  movel([0.238520, -0.777638, -2.781210, -1.153541, 1.570796, 1.809316],accel_mss,speed_ms,0,blend_radius_m)
  movel([0.239014, -0.778562, -2.781058, -1.152769, 1.570796, 1.809811],accel_mss,speed_ms,0,blend_radius_m)
  movel([0.239003, -0.779791, -2.780855, -1.151743, 1.570796, 1.809799],accel_mss,speed_ms,0,blend_radius_m)
  movel([0.238262, -0.781308, -2.780604, -1.150477, 1.570796, 1.809059],accel_mss,speed_ms,0,blend_radius_m)
  movel([0.237067, -0.782563, -2.780395, -1.149431, 1.570796, 1.807864],accel_mss,speed_ms,0,blend_radius_m)
  movel([0.235771, -0.783294, -2.780273, -1.148822, 1.570796, 1.806567],accel_mss,speed_ms,0,blend_radius_m)
  movel([0.234495, -0.783612, -2.780219, -1.148557, 1.570796, 1.805291],accel_mss,speed_ms,0,blend_radius_m)
  movel([0.233364, -0.783640, -2.780215, -1.148534, 1.570796, 1.804160],accel_mss,speed_ms,0,blend_radius_m)
  movel([0.227228, -0.782889, -2.780340, -1.149160, 1.570796, 1.798025],accel_mss,speed_ms,0,blend_radius_m)
  movel([0.221349, -0.781729, -2.780534, -1.150126, 1.570796, 1.792145],accel_mss,speed_ms,0,blend_radius_m)
  movel([0.215730, -0.780164, -2.780794, -1.151432, 1.570796, 1.786526],accel_mss,speed_ms,0,blend_radius_m)
  movel([0.210389, -0.778185, -2.781120, -1.153084, 1.570796, 1.781185],accel_mss,speed_ms,0,blend_radius_m)
  movel([0.208538, -0.777277, -2.781269, -1.153843, 1.570796, 1.779334],accel_mss,speed_ms,0,blend_radius_m)
  movel([0.207075, -0.775893, -2.781496, -1.155000, 1.570796, 1.777871],accel_mss,speed_ms,0,blend_radius_m)
  movel([0.206532, -0.774726, -2.781686, -1.155977, 1.570796, 1.777328],accel_mss,speed_ms,0,blend_radius_m)
  movel([0.206197, -0.773361, -2.781908, -1.157121, 1.570796, 1.776993],accel_mss,speed_ms,0,blend_radius_m)
  movel([0.205895, -0.770284, -2.782404, -1.159701, 1.570796, 1.776692],accel_mss,speed_ms,0,blend_radius_m)
  movel([0.206072, -0.758256, -2.784298, -1.169835, 1.570796, 1.776868],accel_mss,speed_ms,0,blend_radius_m)
  movel([0.205767, -0.755116, -2.784781, -1.172493, 1.570796, 1.776563],accel_mss,speed_ms,0,blend_radius_m)
  movel([0.205061, -0.752630, -2.785159, -1.174600, 1.570796, 1.775857],accel_mss,speed_ms,0,blend_radius_m)
  movel([0.204513, -0.751748, -2.785293, -1.175348, 1.570796, 1.775309],accel_mss,speed_ms,0,blend_radius_m)
  movel([0.203813, -0.751162, -2.785382, -1.175845, 1.570796, 1.774609],accel_mss,speed_ms,0,blend_radius_m)
  movel([0.202946, -0.750924, -2.785418, -1.176048, 1.570796, 1.773742],accel_mss,speed_ms,0,blend_radius_m)
  movel([0.201896, -0.751069, -2.785396, -1.175924, 1.570796, 1.772693],accel_mss,speed_ms,0,blend_radius_m)
  movel([0.199844, -0.751927, -2.785266, -1.175196, 1.570796, 1.770640],accel_mss,speed_ms,0,blend_radius_m)
  movel([0.198900, -0.752216, -2.785222, -1.174950, 1.570796, 1.769696],accel_mss,speed_ms,0,blend_radius_m)
  movel([0.198186, -0.752114, -2.785238, -1.175037, 1.570796, 1.768982],accel_mss,speed_ms,0,blend_radius_m)
  movel([0.197823, -0.751113, -2.785389, -1.175887, 1.570796, 1.768619],accel_mss,speed_ms,0,blend_radius_m)
  movel([0.198037, -0.749591, -2.785618, -1.177180, 1.570796, 1.768834],accel_mss,speed_ms,0,blend_radius_m)
  movel([0.198952, -0.744572, -2.786366, -1.181452, 1.570796, 1.769748],accel_mss,speed_ms,0,blend_radius_m)
  movel([0.199542, -0.739772, -2.787069, -1.185548, 1.570796, 1.770338],accel_mss,speed_ms,0,blend_radius_m)
  movel([0.199909, -0.730710, -2.788367, -1.193312, 1.570796, 1.770705],accel_mss,speed_ms,0,blend_radius_m)
  movel([0.199495, -0.722125, -2.789560, -1.200704, 1.570796, 1.770291],accel_mss,speed_ms,0,blend_radius_m)
  movel([0.198653, -0.713738, -2.790692, -1.207959, 1.570796, 1.769449],accel_mss,speed_ms,0,blend_radius_m)
  speed_ms = 0.005
  movel([0.198653, -0.707172, -2.784094, -1.221123, 1.570796, 1.769449],accel_mss,speed_ms,0,blend_radius_m)
  speed_ms = 0.040
  movel([0.192703, -0.724050, -2.781792, -1.206547, 1.570796, 1.763499],accel_mss,speed_ms,0,blend_radius_m)
  speed_ms = 0.005
  movel([0.192703, -0.730831, -2.788350, -1.193208, 1.570796, 1.763499],accel_mss,speed_ms,0,blend_radius_m)
  speed_ms = 0.025
  movel([0.189482, -0.741949, -2.786751, -1.183689, 1.570796, 1.760279],accel_mss,speed_ms,0,blend_radius_m)
  movel([0.187584, -0.747603, -2.785916, -1.178870, 1.570796, 1.758381],accel_mss,speed_ms,0,blend_radius_m)
  movel([0.185510, -0.753297, -2.785058, -1.174034, 1.570796, 1.756306],accel_mss,speed_ms,0,blend_radius_m)
  movel([0.183050, -0.752490, -2.785181, -1.174719, 1.570796, 1.753846],accel_mss,speed_ms,0,blend_radius_m)
  movel([0.182585, -0.752423, -2.785191, -1.174775, 1.570796, 1.753381],accel_mss,speed_ms,0,blend_radius_m)
  movel([0.182001, -0.752685, -2.785151, -1.174553, 1.570796, 1.752798],accel_mss,speed_ms,0,blend_radius_m)
  movel([0.181431, -0.753357, -2.785049, -1.173983, 1.570796, 1.752227],accel_mss,speed_ms,0,blend_radius_m)
  movel([0.181021, -0.754135, -2.784931, -1.173324, 1.570796, 1.751817],accel_mss,speed_ms,0,blend_radius_m)
  movel([0.178486, -0.758934, -2.784193, -1.169262, 1.570796, 1.749283],accel_mss,speed_ms,0,blend_radius_m)
  movel([0.175445, -0.763691, -2.783451, -1.165247, 1.570796, 1.746242],accel_mss,speed_ms,0,blend_radius_m)
  movel([0.174614, -0.764748, -2.783285, -1.164356, 1.570796, 1.745410],accel_mss,speed_ms,0,blend_radius_m)
  movel([0.173739, -0.765391, -2.783183, -1.163814, 1.570796, 1.744535],accel_mss,speed_ms,0,blend_radius_m)
  movel([0.173247, -0.765240, -2.783207, -1.163942, 1.570796, 1.744044],accel_mss,speed_ms,0,blend_radius_m)
  movel([0.173079, -0.764663, -2.783298, -1.164428, 1.570796, 1.743875],accel_mss,speed_ms,0,blend_radius_m)
  movel([0.172930, -0.760434, -2.783961, -1.167994, 1.570796, 1.743726],accel_mss,speed_ms,0,blend_radius_m)
  movel([0.173553, -0.755646, -2.784700, -1.172043, 1.570796, 1.744349],accel_mss,speed_ms,0,blend_radius_m)
  speed_ms = 0.005
  movel([0.173553, -0.748568, -2.778205, -1.185616, 1.570796, 1.744349],accel_mss,speed_ms,0,blend_radius_m)
  speed_ms = 0.040
  movel([0.180746, -0.753780, -2.777404, -1.181204, 1.570796, 1.751543],accel_mss,speed_ms,0,blend_radius_m)
  speed_ms = 0.005
  movel([0.180746, -0.760919, -2.783885, -1.167585, 1.570796, 1.751543],accel_mss,speed_ms,0,blend_radius_m)
  speed_ms = 0.025
  movel([0.179875, -0.767925, -2.782781, -1.161683, 1.570796, 1.750672],accel_mss,speed_ms,0,blend_radius_m)
  movel([0.179084, -0.771629, -2.782188, -1.158572, 1.570796, 1.749880],accel_mss,speed_ms,0,blend_radius_m)
  movel([0.176839, -0.779327, -2.780932, -1.152130, 1.570796, 1.747635],accel_mss,speed_ms,0,blend_radius_m)
  movel([0.175396, -0.783288, -2.780274, -1.148827, 1.570796, 1.746192],accel_mss,speed_ms,0,blend_radius_m)
  movel([0.171908, -0.791341, -2.778911, -1.142138, 1.570796, 1.742704],accel_mss,speed_ms,0,blend_radius_m)
  movel([0.172377, -0.788931, -2.779322, -1.144136, 1.570796, 1.743174],accel_mss,speed_ms,0,blend_radius_m)
  movel([0.172203, -0.786949, -2.779658, -1.145782, 1.570796, 1.742999],accel_mss,speed_ms,0,blend_radius_m)
  movel([0.171413, -0.785526, -2.779898, -1.146964, 1.570796, 1.742209],accel_mss,speed_ms,0,blend_radius_m)
  movel([0.170034, -0.784796, -2.780021, -1.147572, 1.570796, 1.740831],accel_mss,speed_ms,0,blend_radius_m)
  speed_ms = 0.005
  movel([0.170034, -0.777395, -2.773605, -1.161389, 1.570796, 1.740831],accel_mss,speed_ms,0,blend_radius_m)
  speed_ms = 0.040
  movel([0.144449, -0.795994, -2.770410, -1.145985, 1.570796, 1.715246],accel_mss,speed_ms,0,blend_radius_m)
  speed_ms = 0.005
  movel([0.144449, -0.803590, -2.776772, -1.132027, 1.570796, 1.715246],accel_mss,speed_ms,0,blend_radius_m)
  speed_ms = 0.025
  movel([0.140306, -0.809331, -2.775742, -1.127316, 1.570796, 1.711102],accel_mss,speed_ms,0,blend_radius_m)
  movel([0.135816, -0.814795, -2.774745, -1.122849, 1.570796, 1.706612],accel_mss,speed_ms,0,blend_radius_m)
  movel([0.131062, -0.819901, -2.773799, -1.118689, 1.570796, 1.701858],accel_mss,speed_ms,0,blend_radius_m)
  movel([0.126121, -0.824563, -2.772923, -1.114904, 1.570796, 1.696917],accel_mss,speed_ms,0,blend_radius_m)
  movel([0.127219, -0.822105, -2.773386, -1.116898, 1.570796, 1.698016],accel_mss,speed_ms,0,blend_radius_m)
  movel([0.127994, -0.819853, -2.773808, -1.118728, 1.570796, 1.698790],accel_mss,speed_ms,0,blend_radius_m)
  movel([0.128392, -0.818004, -2.774152, -1.120233, 1.570796, 1.699188],accel_mss,speed_ms,0,blend_radius_m)
  movel([0.128362, -0.816754, -2.774384, -1.121251, 1.570796, 1.699159],accel_mss,speed_ms,0,blend_radius_m)
  movel([0.127847, -0.816316, -2.774465, -1.121608, 1.570796, 1.698643],accel_mss,speed_ms,0,blend_radius_m)
  movel([0.127395, -0.816460, -2.774438, -1.121491, 1.570796, 1.698191],accel_mss,speed_ms,0,blend_radius_m)
  movel([0.126795, -0.816881, -2.774360, -1.121147, 1.570796, 1.697592],accel_mss,speed_ms,0,blend_radius_m)
  movel([0.125163, -0.818650, -2.774032, -1.119707, 1.570796, 1.695960],accel_mss,speed_ms,0,blend_radius_m)
  movel([0.121164, -0.824312, -2.772970, -1.115107, 1.570796, 1.691961],accel_mss,speed_ms,0,blend_radius_m)
  movel([0.119283, -0.826786, -2.772500, -1.113103, 1.570796, 1.690079],accel_mss,speed_ms,0,blend_radius_m)
  movel([0.115192, -0.831505, -2.771595, -1.109289, 1.570796, 1.685989],accel_mss,speed_ms,0,blend_radius_m)
  movel([0.113032, -0.833691, -2.771171, -1.107526, 1.570796, 1.683829],accel_mss,speed_ms,0,blend_radius_m)
  movel([0.110826, -0.835714, -2.770777, -1.105898, 1.570796, 1.681622],accel_mss,speed_ms,0,blend_radius_m)
  movel([0.108596, -0.837553, -2.770416, -1.104420, 1.570796, 1.679392],accel_mss,speed_ms,0,blend_radius_m)
  movel([0.106371, -0.839163, -2.770099, -1.103127, 1.570796, 1.677167],accel_mss,speed_ms,0,blend_radius_m)
  movel([0.108926, -0.835167, -2.770884, -1.106338, 1.570796, 1.679722],accel_mss,speed_ms,0,blend_radius_m)
  movel([0.111408, -0.831132, -2.771667, -1.109590, 1.570796, 1.682204],accel_mss,speed_ms,0,blend_radius_m)
  movel([0.112472, -0.828577, -2.772158, -1.111654, 1.570796, 1.683268],accel_mss,speed_ms,0,blend_radius_m)
  movel([0.112976, -0.826234, -2.772605, -1.113550, 1.570796, 1.683773],accel_mss,speed_ms,0,blend_radius_m)
  movel([0.112833, -0.825536, -2.772738, -1.114115, 1.570796, 1.683630],accel_mss,speed_ms,0,blend_radius_m)
  movel([0.112322, -0.825368, -2.772770, -1.114251, 1.570796, 1.683118],accel_mss,speed_ms,0,blend_radius_m)
  movel([0.111378, -0.825886, -2.772672, -1.113832, 1.570796, 1.682174],accel_mss,speed_ms,0,blend_radius_m)
  movel([0.109924, -0.827249, -2.772412, -1.112728, 1.570796, 1.680720],accel_mss,speed_ms,0,blend_radius_m)
  movel([0.102400, -0.835431, -2.770832, -1.106126, 1.570796, 1.673197],accel_mss,speed_ms,0,blend_radius_m)
  movel([0.098589, -0.839089, -2.770114, -1.103186, 1.570796, 1.669385],accel_mss,speed_ms,0,blend_radius_m)
  movel([0.096654, -0.840643, -2.769806, -1.101939, 1.570796, 1.667451],accel_mss,speed_ms,0,blend_radius_m)
  movel([0.094689, -0.841956, -2.769545, -1.100887, 1.570796, 1.665485],accel_mss,speed_ms,0,blend_radius_m)
  speed_ms = 0.005
  movel([0.094689, -0.834001, -2.763299, -1.115089, 1.570796, 1.665485],accel_mss,speed_ms,0,blend_radius_m)
  speed_ms = 0.040
  movel([0.128026, -0.781141, -2.772976, -1.158272, 1.570796, 1.698822],accel_mss,speed_ms,0,blend_radius_m)
  speed_ms = 0.005
  movel([0.128026, -0.788583, -2.779381, -1.144425, 1.570796, 1.698822],accel_mss,speed_ms,0,blend_radius_m)
  speed_ms = 0.025
  movel([0.127894, -0.785887, -2.779837, -1.146664, 1.570796, 1.698691],accel_mss,speed_ms,0,blend_radius_m)
  movel([0.128371, -0.782803, -2.780355, -1.149231, 1.570796, 1.699168],accel_mss,speed_ms,0,blend_radius_m)
  movel([0.129395, -0.779405, -2.780919, -1.152065, 1.570796, 1.700191],accel_mss,speed_ms,0,blend_radius_m)
  movel([0.130900, -0.775786, -2.781513, -1.155090, 1.570796, 1.701697],accel_mss,speed_ms,0,blend_radius_m)
  movel([0.132838, -0.772016, -2.782125, -1.158247, 1.570796, 1.703635],accel_mss,speed_ms,0,blend_radius_m)
  movel([0.135137, -0.768197, -2.782738, -1.161454, 1.570796, 1.705933],accel_mss,speed_ms,0,blend_radius_m)
  movel([0.137743, -0.764400, -2.783340, -1.164649, 1.570796, 1.708540],accel_mss,speed_ms,0,blend_radius_m)
  movel([0.140583, -0.760728, -2.783915, -1.167746, 1.570796, 1.711379],accel_mss,speed_ms,0,blend_radius_m)
  movel([0.144308, -0.756402, -2.784584, -1.171403, 1.570796, 1.715105],accel_mss,speed_ms,0,blend_radius_m)
  movel([0.151976, -0.747852, -2.785879, -1.178659, 1.570796, 1.722772],accel_mss,speed_ms,0,blend_radius_m)
  movel([0.155648, -0.743371, -2.786543, -1.182475, 1.570796, 1.726445],accel_mss,speed_ms,0,blend_radius_m)
  movel([0.158985, -0.738544, -2.787247, -1.186598, 1.570796, 1.729782],accel_mss,speed_ms,0,blend_radius_m)
  movel([0.160417, -0.736070, -2.787604, -1.188715, 1.570796, 1.731214],accel_mss,speed_ms,0,blend_radius_m)
  movel([0.161621, -0.733642, -2.787951, -1.190796, 1.570796, 1.732417],accel_mss,speed_ms,0,blend_radius_m)
  movel([0.162542, -0.731323, -2.788280, -1.192786, 1.570796, 1.733339],accel_mss,speed_ms,0,blend_radius_m)
  movel([0.163134, -0.729175, -2.788583, -1.194631, 1.570796, 1.733930],accel_mss,speed_ms,0,blend_radius_m)
  movel([0.163330, -0.727280, -2.788848, -1.196261, 1.570796, 1.734126],accel_mss,speed_ms,0,blend_radius_m)
  movel([0.163076, -0.725704, -2.789067, -1.197618, 1.570796, 1.733872],accel_mss,speed_ms,0,blend_radius_m)
  speed_ms = 0.005
  movel([0.163076, -0.718987, -2.782497, -1.210906, 1.570796, 1.733872],accel_mss,speed_ms,0,blend_radius_m)
  speed_ms = 0.040
  movel([0.160050, -0.707154, -2.784096, -1.221139, 1.570796, 1.730846],accel_mss,speed_ms,0,blend_radius_m)
  speed_ms = 0.005
  movel([0.160050, -0.713719, -2.790695, -1.207975, 1.570796, 1.730846],accel_mss,speed_ms,0,blend_radius_m)
  speed_ms = 0.025
  movel([0.157424, -0.725682, -2.789070, -1.197637, 1.570796, 1.728221],accel_mss,speed_ms,0,blend_radius_m)
  movel([0.156311, -0.728566, -2.788668, -1.195155, 1.570796, 1.727108],accel_mss,speed_ms,0,blend_radius_m)
  movel([0.154500, -0.731547, -2.788249, -1.192593, 1.570796, 1.725296],accel_mss,speed_ms,0,blend_radius_m)
  movel([0.152223, -0.734414, -2.787841, -1.190134, 1.570796, 1.723019],accel_mss,speed_ms,0,blend_radius_m)
  movel([0.144460, -0.743032, -2.786593, -1.182764, 1.570796, 1.715257],accel_mss,speed_ms,0,blend_radius_m)
  movel([0.141887, -0.746260, -2.786116, -1.180013, 1.570796, 1.712683],accel_mss,speed_ms,0,blend_radius_m)
  movel([0.139486, -0.749568, -2.785622, -1.177199, 1.570796, 1.710282],accel_mss,speed_ms,0,blend_radius_m)
  movel([0.137275, -0.752916, -2.785116, -1.174357, 1.570796, 1.708071],accel_mss,speed_ms,0,blend_radius_m)
  movel([0.135464, -0.756183, -2.784617, -1.171588, 1.570796, 1.706261],accel_mss,speed_ms,0,blend_radius_m)
  movel([0.133979, -0.759398, -2.784121, -1.168869, 1.570796, 1.704776],accel_mss,speed_ms,0,blend_radius_m)
  movel([0.132528, -0.762585, -2.783625, -1.166179, 1.570796, 1.703325],accel_mss,speed_ms,0,blend_radius_m)
  movel([0.130825, -0.765773, -2.783123, -1.163493, 1.570796, 1.701621],accel_mss,speed_ms,0,blend_radius_m)
  movel([0.128528, -0.761127, -2.783853, -1.167409, 1.570796, 1.699324],accel_mss,speed_ms,0,blend_radius_m)
  movel([0.128585, -0.759365, -2.784127, -1.168898, 1.570796, 1.699381],accel_mss,speed_ms,0,blend_radius_m)
  movel([0.128955, -0.757448, -2.784423, -1.170518, 1.570796, 1.699752],accel_mss,speed_ms,0,blend_radius_m)
  movel([0.129638, -0.755372, -2.784742, -1.172275, 1.570796, 1.700435],accel_mss,speed_ms,0,blend_radius_m)
  movel([0.130651, -0.753118, -2.785085, -1.174186, 1.570796, 1.701447],accel_mss,speed_ms,0,blend_radius_m)
  movel([0.132666, -0.749871, -2.785576, -1.176942, 1.570796, 1.703462],accel_mss,speed_ms,0,blend_radius_m)
  movel([0.135700, -0.745820, -2.786181, -1.180388, 1.570796, 1.706497],accel_mss,speed_ms,0,blend_radius_m)
  movel([0.143277, -0.736531, -2.787538, -1.188320, 1.570796, 1.714073],accel_mss,speed_ms,0,blend_radius_m)
  movel([0.147031, -0.731929, -2.788195, -1.192265, 1.570796, 1.717828],accel_mss,speed_ms,0,blend_radius_m)
  movel([0.150221, -0.727782, -2.788778, -1.195829, 1.570796, 1.721017],accel_mss,speed_ms,0,blend_radius_m)
  movel([0.152429, -0.724431, -2.789243, -1.198715, 1.570796, 1.723225],accel_mss,speed_ms,0,blend_radius_m)
  movel([0.153036, -0.723152, -2.789419, -1.199818, 1.570796, 1.723833],accel_mss,speed_ms,0,blend_radius_m)
  movel([0.153239, -0.722197, -2.789550, -1.200642, 1.570796, 1.724035],accel_mss,speed_ms,0,blend_radius_m)
  speed_ms = 0.005
  movel([0.153239, -0.715524, -2.782972, -1.213894, 1.570796, 1.724035],accel_mss,speed_ms,0,blend_radius_m)
  speed_ms = 0.040
  movel([0.137879, -0.720219, -2.782326, -1.209843, 1.570796, 1.708675],accel_mss,speed_ms,0,blend_radius_m)
  speed_ms = 0.005
  movel([0.137879, -0.726952, -2.788893, -1.196543, 1.570796, 1.708675],accel_mss,speed_ms,0,blend_radius_m)
  speed_ms = 0.025
  movel([0.136395, -0.727386, -2.788833, -1.196170, 1.570796, 1.707191],accel_mss,speed_ms,0,blend_radius_m)
  movel([0.135134, -0.727419, -2.788828, -1.196142, 1.570796, 1.705931],accel_mss,speed_ms,0,blend_radius_m)
  movel([0.133190, -0.726532, -2.788952, -1.196905, 1.570796, 1.703986],accel_mss,speed_ms,0,blend_radius_m)
  movel([0.131847, -0.724748, -2.789199, -1.198441, 1.570796, 1.702644],accel_mss,speed_ms,0,blend_radius_m)
  movel([0.130926, -0.722510, -2.789507, -1.200371, 1.570796, 1.701722],accel_mss,speed_ms,0,blend_radius_m)
  movel([0.130785, -0.721530, -2.789642, -1.201218, 1.570796, 1.701582],accel_mss,speed_ms,0,blend_radius_m)
  movel([0.131601, -0.719398, -2.789932, -1.203059, 1.570796, 1.702397],accel_mss,speed_ms,0,blend_radius_m)
  movel([0.134610, -0.713129, -2.790773, -1.208487, 1.570796, 1.705407],accel_mss,speed_ms,0,blend_radius_m)
  movel([0.140137, -0.700606, -2.792400, -1.219383, 1.570796, 1.710933],accel_mss,speed_ms,0,blend_radius_m)
  movel([0.142639, -0.694384, -2.793181, -1.224825, 1.570796, 1.713435],accel_mss,speed_ms,0,blend_radius_m)
  speed_ms = 0.005
  movel([0.142639, -0.688072, -2.786538, -1.237779, 1.570796, 1.713435],accel_mss,speed_ms,0,blend_radius_m)
  speed_ms = 0.040
  movel([0.132933, -0.695886, -2.785558, -1.230945, 1.570796, 1.703729],accel_mss,speed_ms,0,blend_radius_m)
  speed_ms = 0.005
  movel([0.132933, -0.702302, -2.792184, -1.217903, 1.570796, 1.703729],accel_mss,speed_ms,0,blend_radius_m)
  speed_ms = 0.025
  movel([0.131774, -0.705905, -2.791720, -1.214763, 1.570796, 1.702571],accel_mss,speed_ms,0,blend_radius_m)
  movel([0.130233, -0.709651, -2.791232, -1.211506, 1.570796, 1.701029],accel_mss,speed_ms,0,blend_radius_m)
  movel([0.128199, -0.713401, -2.790737, -1.208251, 1.570796, 1.698995],accel_mss,speed_ms,0,blend_radius_m)
  movel([0.126962, -0.715242, -2.790492, -1.206655, 1.570796, 1.697758],accel_mss,speed_ms,0,blend_radius_m)
  movel([0.124214, -0.718795, -2.790014, -1.203580, 1.570796, 1.695010],accel_mss,speed_ms,0,blend_radius_m)
  movel([0.123618, -0.720283, -2.789812, -1.202294, 1.570796, 1.694414],accel_mss,speed_ms,0,blend_radius_m)
  movel([0.120317, -0.731224, -2.788294, -1.192871, 1.570796, 1.691113],accel_mss,speed_ms,0,blend_radius_m)
  movel([0.120030, -0.732265, -2.788147, -1.191977, 1.570796, 1.690826],accel_mss,speed_ms,0,blend_radius_m)
  movel([0.120015, -0.733114, -2.788027, -1.191249, 1.570796, 1.690811],accel_mss,speed_ms,0,blend_radius_m)
  movel([0.120743, -0.733613, -2.787955, -1.190820, 1.570796, 1.691539],accel_mss,speed_ms,0,blend_radius_m)
  movel([0.121930, -0.733493, -2.787972, -1.190923, 1.570796, 1.692726],accel_mss,speed_ms,0,blend_radius_m)
  movel([0.125409, -0.732988, -2.788044, -1.191356, 1.570796, 1.696206],accel_mss,speed_ms,0,blend_radius_m)
  movel([0.128620, -0.732965, -2.788048, -1.191376, 1.570796, 1.699416],accel_mss,speed_ms,0,blend_radius_m)
  movel([0.131341, -0.733654, -2.787950, -1.190785, 1.570796, 1.702138],accel_mss,speed_ms,0,blend_radius_m)
  movel([0.133335, -0.735302, -2.787714, -1.189373, 1.570796, 1.704131],accel_mss,speed_ms,0,blend_radius_m)
  speed_ms = 0.005
  movel([0.133335, -0.728466, -2.781168, -1.202756, 1.570796, 1.704131],accel_mss,speed_ms,0,blend_radius_m)
  speed_ms = 0.040
  movel([0.124946, -0.756050, -2.777052, -1.179288, 1.570796, 1.695742],accel_mss,speed_ms,0,blend_radius_m)
  speed_ms = 0.005
  movel([0.124946, -0.763214, -2.783526, -1.165648, 1.570796, 1.695742],accel_mss,speed_ms,0,blend_radius_m)
  speed_ms = 0.025
  movel([0.124279, -0.763945, -2.783411, -1.165033, 1.570796, 1.695076],accel_mss,speed_ms,0,blend_radius_m)
  movel([0.123694, -0.764818, -2.783274, -1.164297, 1.570796, 1.694491],accel_mss,speed_ms,0,blend_radius_m)
  movel([0.121456, -0.769175, -2.782582, -1.160632, 1.570796, 1.692253],accel_mss,speed_ms,0,blend_radius_m)
  movel([0.121055, -0.769619, -2.782511, -1.160259, 1.570796, 1.691851],accel_mss,speed_ms,0,blend_radius_m)
  movel([0.120432, -0.769904, -2.782465, -1.160020, 1.570796, 1.691229],accel_mss,speed_ms,0,blend_radius_m)
  movel([0.119925, -0.769768, -2.782487, -1.160134, 1.570796, 1.690722],accel_mss,speed_ms,0,blend_radius_m)
  movel([0.119237, -0.768645, -2.782667, -1.161078, 1.570796, 1.690033],accel_mss,speed_ms,0,blend_radius_m)
  movel([0.118835, -0.765855, -2.783110, -1.163424, 1.570796, 1.689631],accel_mss,speed_ms,0,blend_radius_m)
  movel([0.119383, -0.762634, -2.783617, -1.166137, 1.570796, 1.690179],accel_mss,speed_ms,0,blend_radius_m)
  movel([0.120418, -0.759122, -2.784164, -1.169102, 1.570796, 1.691215],accel_mss,speed_ms,0,blend_radius_m)
  movel([0.121709, -0.755540, -2.784716, -1.172133, 1.570796, 1.692506],accel_mss,speed_ms,0,blend_radius_m)
  movel([0.123298, -0.751966, -2.785260, -1.175163, 1.570796, 1.694094],accel_mss,speed_ms,0,blend_radius_m)
  movel([0.125173, -0.748402, -2.785796, -1.178190, 1.570796, 1.695969],accel_mss,speed_ms,0,blend_radius_m)
  movel([0.127322, -0.744851, -2.786324, -1.181213, 1.570796, 1.698119],accel_mss,speed_ms,0,blend_radius_m)
  movel([0.129739, -0.741309, -2.786845, -1.184235, 1.570796, 1.700535],accel_mss,speed_ms,0,blend_radius_m)
  movel([0.132404, -0.737785, -2.787357, -1.187247, 1.570796, 1.703200],accel_mss,speed_ms,0,blend_radius_m)
  movel([0.135317, -0.734268, -2.787862, -1.190259, 1.570796, 1.706113],accel_mss,speed_ms,0,blend_radius_m)
  movel([0.138458, -0.730769, -2.788359, -1.193261, 1.570796, 1.709254],accel_mss,speed_ms,0,blend_radius_m)
  movel([0.142773, -0.725595, -2.789082, -1.197712, 1.570796, 1.713570],accel_mss,speed_ms,0,blend_radius_m)
  movel([0.147235, -0.719614, -2.789903, -1.202872, 1.570796, 1.718031],accel_mss,speed_ms,0,blend_radius_m)
  movel([0.152015, -0.712739, -2.790825, -1.208825, 1.570796, 1.722812],accel_mss,speed_ms,0,blend_radius_m)
  speed_ms = 0.005
  movel([0.152015, -0.706186, -2.784224, -1.221979, 1.570796, 1.722812],accel_mss,speed_ms,0,blend_radius_m)
  speed_ms = 0.040
  movel([0.147515, -0.708228, -2.783953, -1.220207, 1.570796, 1.718311],accel_mss,speed_ms,0,blend_radius_m)
  speed_ms = 0.005
  movel([0.147515, -0.714808, -2.790550, -1.207031, 1.570796, 1.718311],accel_mss,speed_ms,0,blend_radius_m)
  speed_ms = 0.025
  movel([0.150955, -0.705951, -2.791714, -1.214723, 1.570796, 1.721751],accel_mss,speed_ms,0,blend_radius_m)
  movel([0.154901, -0.696855, -2.792873, -1.222662, 1.570796, 1.725698],accel_mss,speed_ms,0,blend_radius_m)
  movel([0.157180, -0.692234, -2.793447, -1.226708, 1.570796, 1.727976],accel_mss,speed_ms,0,blend_radius_m)
  movel([0.159708, -0.687580, -2.794015, -1.230794, 1.570796, 1.730504],accel_mss,speed_ms,0,blend_radius_m)
  movel([0.162546, -0.682891, -2.794578, -1.234920, 1.570796, 1.733342],accel_mss,speed_ms,0,blend_radius_m)
  movel([0.165720, -0.678193, -2.795132, -1.239064, 1.570796, 1.736517],accel_mss,speed_ms,0,blend_radius_m)
  movel([0.174701, -0.666260, -2.796496, -1.249633, 1.570796, 1.745498],accel_mss,speed_ms,0,blend_radius_m)
  movel([0.178567, -0.660821, -2.797097, -1.254472, 1.570796, 1.749363],accel_mss,speed_ms,0,blend_radius_m)
  movel([0.180369, -0.658058, -2.797397, -1.256934, 1.570796, 1.751165],accel_mss,speed_ms,0,blend_radius_m)
  movel([0.181974, -0.655275, -2.797696, -1.259418, 1.570796, 1.752770],accel_mss,speed_ms,0,blend_radius_m)
  movel([0.185372, -0.647161, -2.798550, -1.266679, 1.570796, 1.756168],accel_mss,speed_ms,0,blend_radius_m)
  speed_ms = 0.005
  movel([0.185372, -0.641516, -2.791809, -1.279065, 1.570796, 1.756168],accel_mss,speed_ms,0,blend_radius_m)
  speed_ms = 0.040
  movel([0.193729, -0.622779, -2.793665, -1.295945, 1.570796, 1.764526],accel_mss,speed_ms,0,blend_radius_m)
  speed_ms = 0.005
  movel([0.193729, -0.628139, -2.800441, -1.283810, 1.570796, 1.764526],accel_mss,speed_ms,0,blend_radius_m)
  speed_ms = 0.025
  movel([0.196333, -0.621490, -2.801066, -1.289833, 1.570796, 1.767130],accel_mss,speed_ms,0,blend_radius_m)
  movel([0.198154, -0.618053, -2.801382, -1.292954, 1.570796, 1.768950],accel_mss,speed_ms,0,blend_radius_m)
  movel([0.200526, -0.614603, -2.801695, -1.296091, 1.570796, 1.771322],accel_mss,speed_ms,0,blend_radius_m)
  movel([0.202505, -0.612299, -2.801901, -1.298189, 1.570796, 1.773301],accel_mss,speed_ms,0,blend_radius_m)
  movel([0.204614, -0.610164, -2.802090, -1.300135, 1.570796, 1.775410],accel_mss,speed_ms,0,blend_radius_m)
  movel([0.209001, -0.606162, -2.802439, -1.303789, 1.570796, 1.779798],accel_mss,speed_ms,0,blend_radius_m)
  movel([0.212909, -0.602297, -2.802770, -1.307322, 1.570796, 1.783705],accel_mss,speed_ms,0,blend_radius_m)
  movel([0.215989, -0.598561, -2.803084, -1.310744, 1.570796, 1.786785],accel_mss,speed_ms,0,blend_radius_m)
  movel([0.221767, -0.590075, -2.803777, -1.318537, 1.570796, 1.792563],accel_mss,speed_ms,0,blend_radius_m)
  movel([0.223037, -0.588369, -2.803913, -1.320107, 1.570796, 1.793834],accel_mss,speed_ms,0,blend_radius_m)
  movel([0.224449, -0.586785, -2.804038, -1.321566, 1.570796, 1.795245],accel_mss,speed_ms,0,blend_radius_m)
  movel([0.227568, -0.583894, -2.804264, -1.324231, 1.570796, 1.798364],accel_mss,speed_ms,0,blend_radius_m)
  movel([0.233995, -0.578551, -2.804672, -1.329165, 1.570796, 1.804791],accel_mss,speed_ms,0,blend_radius_m)
  movel([0.240772, -0.572320, -2.805135, -1.334934, 1.570796, 1.811568],accel_mss,speed_ms,0,blend_radius_m)
  movel([0.244115, -0.568952, -2.805378, -1.338059, 1.570796, 1.814911],accel_mss,speed_ms,0,blend_radius_m)
  movel([0.247325, -0.565306, -2.805637, -1.341446, 1.570796, 1.818121],accel_mss,speed_ms,0,blend_radius_m)
  movel([0.249641, -0.562122, -2.805859, -1.344408, 1.570796, 1.820438],accel_mss,speed_ms,0,blend_radius_m)
  movel([0.251409, -0.558950, -2.806075, -1.347363, 1.570796, 1.822205],accel_mss,speed_ms,0,blend_radius_m)
  movel([0.252187, -0.556399, -2.806247, -1.349743, 1.570796, 1.822983],accel_mss,speed_ms,0,blend_radius_m)
  movel([0.252068, -0.555552, -2.806304, -1.350534, 1.570796, 1.822864],accel_mss,speed_ms,0,blend_radius_m)
  movel([0.251533, -0.555093, -2.806334, -1.350962, 1.570796, 1.822330],accel_mss,speed_ms,0,blend_radius_m)
  movel([0.249691, -0.555064, -2.806336, -1.350989, 1.570796, 1.820487],accel_mss,speed_ms,0,blend_radius_m)
  movel([0.247199, -0.555806, -2.806287, -1.350296, 1.570796, 1.817995],accel_mss,speed_ms,0,blend_radius_m)
  movel([0.244223, -0.557208, -2.806193, -1.348988, 1.570796, 1.815020],accel_mss,speed_ms,0,blend_radius_m)
  movel([0.240967, -0.559117, -2.806064, -1.347208, 1.570796, 1.811764],accel_mss,speed_ms,0,blend_radius_m)
  movel([0.237607, -0.561424, -2.805907, -1.345059, 1.570796, 1.808403],accel_mss,speed_ms,0,blend_radius_m)
  movel([0.234331, -0.563983, -2.805729, -1.342677, 1.570796, 1.805127],accel_mss,speed_ms,0,blend_radius_m)
  movel([0.231319, -0.566673, -2.805541, -1.340176, 1.570796, 1.802115],accel_mss,speed_ms,0,blend_radius_m)
  movel([0.228747, -0.569367, -2.805348, -1.337674, 1.570796, 1.799543],accel_mss,speed_ms,0,blend_radius_m)
  movel([0.225354, -0.573742, -2.805031, -1.333617, 1.570796, 1.796150],accel_mss,speed_ms,0,blend_radius_m)
  movel([0.216091, -0.586999, -2.804021, -1.321368, 1.570796, 1.786887],accel_mss,speed_ms,0,blend_radius_m)
  movel([0.209605, -0.595587, -2.803330, -1.313472, 1.570796, 1.780401],accel_mss,speed_ms,0,blend_radius_m)
  movel([0.203573, -0.602636, -2.802741, -1.307012, 1.570796, 1.774369],accel_mss,speed_ms,0,blend_radius_m)
  movel([0.200581, -0.606065, -2.802447, -1.303877, 1.570796, 1.771378],accel_mss,speed_ms,0,blend_radius_m)
  movel([0.197793, -0.609574, -2.802142, -1.300674, 1.570796, 1.768589],accel_mss,speed_ms,0,blend_radius_m)
  movel([0.195217, -0.613309, -2.801811, -1.297269, 1.570796, 1.766013],accel_mss,speed_ms,0,blend_radius_m)
  movel([0.192956, -0.617013, -2.801477, -1.293898, 1.570796, 1.763753],accel_mss,speed_ms,0,blend_radius_m)
  movel([0.190975, -0.620680, -2.801141, -1.290568, 1.570796, 1.761772],accel_mss,speed_ms,0,blend_radius_m)
  movel([0.189235, -0.624290, -2.800805, -1.287294, 1.570796, 1.760032],accel_mss,speed_ms,0,blend_radius_m)
  movel([0.186322, -0.631317, -2.800135, -1.280937, 1.570796, 1.757118],accel_mss,speed_ms,0,blend_radius_m)
  movel([0.183895, -0.638024, -2.799477, -1.274888, 1.570796, 1.754691],accel_mss,speed_ms,0,blend_radius_m)
  speed_ms = 0.005
  movel([0.183895, -0.632515, -2.792719, -1.287155, 1.570796, 1.754691],accel_mss,speed_ms,0,blend_radius_m)
  speed_ms = 0.040
  movel([0.176152, -0.639775, -2.791987, -1.280627, 1.570796, 1.746948],accel_mss,speed_ms,0,blend_radius_m)
  speed_ms = 0.005
  movel([0.176152, -0.645394, -2.798732, -1.268264, 1.570796, 1.746948],accel_mss,speed_ms,0,blend_radius_m)
  speed_ms = 0.025
  movel([0.180224, -0.634747, -2.799801, -1.277841, 1.570796, 1.751020],accel_mss,speed_ms,0,blend_radius_m)
  movel([0.182120, -0.630206, -2.800243, -1.281940, 1.570796, 1.752916],accel_mss,speed_ms,0,blend_radius_m)
  movel([0.183798, -0.625753, -2.800667, -1.285969, 1.570796, 1.754594],accel_mss,speed_ms,0,blend_radius_m)
  movel([0.184805, -0.622128, -2.801007, -1.289254, 1.570796, 1.755601],accel_mss,speed_ms,0,blend_radius_m)
  movel([0.185326, -0.618806, -2.801313, -1.292269, 1.570796, 1.756122],accel_mss,speed_ms,0,blend_radius_m)
  movel([0.185349, -0.615856, -2.801582, -1.294951, 1.570796, 1.756145],accel_mss,speed_ms,0,blend_radius_m)
  movel([0.184865, -0.613347, -2.801807, -1.297234, 1.570796, 1.755661],accel_mss,speed_ms,0,blend_radius_m)
  movel([0.186494, -0.611974, -2.801930, -1.298485, 1.570796, 1.757290],accel_mss,speed_ms,0,blend_radius_m)
  movel([0.188104, -0.610937, -2.802022, -1.299431, 1.570796, 1.758900],accel_mss,speed_ms,0,blend_radius_m)
  movel([0.191272, -0.609291, -2.802166, -1.300932, 1.570796, 1.762069],accel_mss,speed_ms,0,blend_radius_m)
  movel([0.194593, -0.607312, -2.802339, -1.302738, 1.570796, 1.765389],accel_mss,speed_ms,0,blend_radius_m)
  movel([0.196244, -0.605965, -2.802456, -1.303968, 1.570796, 1.767041],accel_mss,speed_ms,0,blend_radius_m)
  movel([0.197767, -0.604278, -2.802601, -1.305510, 1.570796, 1.768564],accel_mss,speed_ms,0,blend_radius_m)
  movel([0.214731, -0.582487, -2.804372, -1.325529, 1.570796, 1.785527],accel_mss,speed_ms,0,blend_radius_m)
  movel([0.214676, -0.580480, -2.804526, -1.327383, 1.570796, 1.785472],accel_mss,speed_ms,0,blend_radius_m)
  movel([0.213877, -0.579104, -2.804631, -1.328655, 1.570796, 1.784674],accel_mss,speed_ms,0,blend_radius_m)
  movel([0.212377, -0.578432, -2.804681, -1.329276, 1.570796, 1.783174],accel_mss,speed_ms,0,blend_radius_m)
  movel([0.210246, -0.578518, -2.804675, -1.329196, 1.570796, 1.781042],accel_mss,speed_ms,0,blend_radius_m)
  movel([0.214128, -0.575879, -2.804873, -1.331638, 1.570796, 1.784924],accel_mss,speed_ms,0,blend_radius_m)
  movel([0.217788, -0.573955, -2.805015, -1.333419, 1.570796, 1.788584],accel_mss,speed_ms,0,blend_radius_m)
  movel([0.221033, -0.572837, -2.805097, -1.334456, 1.570796, 1.791829],accel_mss,speed_ms,0,blend_radius_m)
  movel([0.223683, -0.572603, -2.805114, -1.334672, 1.570796, 1.794480],accel_mss,speed_ms,0,blend_radius_m)
  speed_ms = 0.005
  movel([0.223683, -0.568129, -2.798249, -1.346011, 1.570796, 1.794480],accel_mss,speed_ms,0,blend_radius_m)
  speed_ms = 0.040
  movel([0.226080, -0.558963, -2.798901, -1.354525, 1.570796, 1.796876],accel_mss,speed_ms,0,blend_radius_m)
  speed_ms = 0.005
  movel([0.226080, -0.563281, -2.805778, -1.343330, 1.570796, 1.796876],accel_mss,speed_ms,0,blend_radius_m)
  speed_ms = 0.025
  movel([0.228138, -0.557951, -2.806143, -1.348295, 1.570796, 1.798934],accel_mss,speed_ms,0,blend_radius_m)
  movel([0.229724, -0.553041, -2.806469, -1.352878, 1.570796, 1.800520],accel_mss,speed_ms,0,blend_radius_m)
  movel([0.230868, -0.548512, -2.806762, -1.357115, 1.570796, 1.801665],accel_mss,speed_ms,0,blend_radius_m)
  movel([0.231595, -0.544322, -2.807026, -1.361041, 1.570796, 1.802391],accel_mss,speed_ms,0,blend_radius_m)
  movel([0.231931, -0.540427, -2.807265, -1.364697, 1.570796, 1.802727],accel_mss,speed_ms,0,blend_radius_m)
  movel([0.231904, -0.536780, -2.807484, -1.368125, 1.570796, 1.802701],accel_mss,speed_ms,0,blend_radius_m)
  movel([0.230885, -0.530050, -2.807875, -1.374465, 1.570796, 1.801682],accel_mss,speed_ms,0,blend_radius_m)
  movel([0.224092, -0.548238, -2.806779, -1.357371, 1.570796, 1.794888],accel_mss,speed_ms,0,blend_radius_m)
  movel([0.224651, -0.546332, -2.806900, -1.359157, 1.570796, 1.795447],accel_mss,speed_ms,0,blend_radius_m)
  movel([0.224852, -0.544671, -2.807004, -1.360714, 1.570796, 1.795649],accel_mss,speed_ms,0,blend_radius_m)
  movel([0.224312, -0.542032, -2.807167, -1.363190, 1.570796, 1.795109],accel_mss,speed_ms,0,blend_radius_m)
  movel([0.222714, -0.540224, -2.807278, -1.364887, 1.570796, 1.793510],accel_mss,speed_ms,0,blend_radius_m)
  movel([0.220333, -0.539136, -2.807343, -1.365909, 1.570796, 1.791129],accel_mss,speed_ms,0,blend_radius_m)
  movel([0.217432, -0.538649, -2.807373, -1.366367, 1.570796, 1.788229],accel_mss,speed_ms,0,blend_radius_m)
  movel([0.214292, -0.538644, -2.807373, -1.366372, 1.570796, 1.785088],accel_mss,speed_ms,0,blend_radius_m)
  movel([0.208391, -0.539580, -2.807317, -1.365493, 1.570796, 1.779188],accel_mss,speed_ms,0,blend_radius_m)
  movel([0.211122, -0.543986, -2.807047, -1.361356, 1.570796, 1.781918],accel_mss,speed_ms,0,blend_radius_m)
  movel([0.211813, -0.546927, -2.806863, -1.358599, 1.570796, 1.782610],accel_mss,speed_ms,0,blend_radius_m)
  movel([0.211526, -0.550446, -2.806638, -1.355305, 1.570796, 1.782322],accel_mss,speed_ms,0,blend_radius_m)
  movel([0.209060, -0.551580, -2.806565, -1.354245, 1.570796, 1.779856],accel_mss,speed_ms,0,blend_radius_m)
  movel([0.206761, -0.552256, -2.806521, -1.353612, 1.570796, 1.777558],accel_mss,speed_ms,0,blend_radius_m)
  movel([0.202396, -0.552864, -2.806481, -1.353044, 1.570796, 1.773192],accel_mss,speed_ms,0,blend_radius_m)
  movel([0.197929, -0.553484, -2.806440, -1.352464, 1.570796, 1.768725],accel_mss,speed_ms,0,blend_radius_m)
  movel([0.195504, -0.554176, -2.806395, -1.351818, 1.570796, 1.766300],accel_mss,speed_ms,0,blend_radius_m)
  movel([0.192883, -0.555309, -2.806320, -1.350760, 1.570796, 1.763679],accel_mss,speed_ms,0,blend_radius_m)
  movel([0.190652, -0.560199, -2.805991, -1.346199, 1.570796, 1.761448],accel_mss,speed_ms,0,blend_radius_m)
  movel([0.189350, -0.564603, -2.805686, -1.342100, 1.570796, 1.760146],accel_mss,speed_ms,0,blend_radius_m)
  movel([0.185745, -0.566570, -2.805548, -1.340271, 1.570796, 1.756542],accel_mss,speed_ms,0,blend_radius_m)
  movel([0.182404, -0.567911, -2.805453, -1.339025, 1.570796, 1.753200],accel_mss,speed_ms,0,blend_radius_m)
  movel([0.179388, -0.568602, -2.805403, -1.338384, 1.570796, 1.750184],accel_mss,speed_ms,0,blend_radius_m)
  movel([0.176782, -0.568621, -2.805402, -1.338366, 1.570796, 1.747579],accel_mss,speed_ms,0,blend_radius_m)
  movel([0.176392, -0.569179, -2.805362, -1.337848, 1.570796, 1.747188],accel_mss,speed_ms,0,blend_radius_m)
  movel([0.173374, -0.575341, -2.804912, -1.332135, 1.570796, 1.744170],accel_mss,speed_ms,0,blend_radius_m)
  movel([0.169984, -0.582867, -2.804343, -1.325179, 1.570796, 1.740781],accel_mss,speed_ms,0,blend_radius_m)
  movel([0.168807, -0.586291, -2.804077, -1.322021, 1.570796, 1.739603],accel_mss,speed_ms,0,blend_radius_m)
  movel([0.168021, -0.589300, -2.803839, -1.319250, 1.570796, 1.738817],accel_mss,speed_ms,0,blend_radius_m)
  movel([0.167144, -0.595092, -2.803371, -1.313927, 1.570796, 1.737940],accel_mss,speed_ms,0,blend_radius_m)
  movel([0.158403, -0.593767, -2.803479, -1.315143, 1.570796, 1.729200],accel_mss,speed_ms,0,blend_radius_m)
  movel([0.157042, -0.597412, -2.803180, -1.311797, 1.570796, 1.727839],accel_mss,speed_ms,0,blend_radius_m)
  movel([0.155985, -0.600919, -2.802886, -1.308583, 1.570796, 1.726781],accel_mss,speed_ms,0,blend_radius_m)
  movel([0.154661, -0.607511, -2.802322, -1.302556, 1.570796, 1.725457],accel_mss,speed_ms,0,blend_radius_m)
  movel([0.154262, -0.613434, -2.801800, -1.297156, 1.570796, 1.725059],accel_mss,speed_ms,0,blend_radius_m)
  movel([0.154695, -0.620188, -2.801187, -1.291014, 1.570796, 1.725492],accel_mss,speed_ms,0,blend_radius_m)
  movel([0.154495, -0.621135, -2.801099, -1.290155, 1.570796, 1.725292],accel_mss,speed_ms,0,blend_radius_m)
  movel([0.154014, -0.622210, -2.800999, -1.289180, 1.570796, 1.724810],accel_mss,speed_ms,0,blend_radius_m)
  movel([0.152932, -0.623706, -2.800860, -1.287824, 1.570796, 1.723728],accel_mss,speed_ms,0,blend_radius_m)
  movel([0.144473, -0.632526, -2.800018, -1.279845, 1.570796, 1.715269],accel_mss,speed_ms,0,blend_radius_m)
  movel([0.140094, -0.636517, -2.799627, -1.276246, 1.570796, 1.710890],accel_mss,speed_ms,0,blend_radius_m)
  movel([0.138438, -0.637671, -2.799512, -1.275206, 1.570796, 1.709235],accel_mss,speed_ms,0,blend_radius_m)
  movel([0.137413, -0.637922, -2.799487, -1.274980, 1.570796, 1.708210],accel_mss,speed_ms,0,blend_radius_m)
  movel([0.141719, -0.639134, -2.799366, -1.273889, 1.570796, 1.712515],accel_mss,speed_ms,0,blend_radius_m)
  movel([0.144168, -0.639301, -2.799349, -1.273738, 1.570796, 1.714964],accel_mss,speed_ms,0,blend_radius_m)
  movel([0.146793, -0.639184, -2.799361, -1.273844, 1.570796, 1.717590],accel_mss,speed_ms,0,blend_radius_m)
  movel([0.139951, -0.648730, -2.798387, -1.265272, 1.570796, 1.710748],accel_mss,speed_ms,0,blend_radius_m)
  movel([0.132855, -0.659158, -2.797278, -1.255953, 1.570796, 1.703651],accel_mss,speed_ms,0,blend_radius_m)
  movel([0.129573, -0.664371, -2.796706, -1.251312, 1.570796, 1.700369],accel_mss,speed_ms,0,blend_radius_m)
  movel([0.126649, -0.669403, -2.796143, -1.246843, 1.570796, 1.697445],accel_mss,speed_ms,0,blend_radius_m)
  movel([0.124224, -0.674136, -2.795603, -1.242650, 1.570796, 1.695020],accel_mss,speed_ms,0,blend_radius_m)
  movel([0.122426, -0.678439, -2.795103, -1.238847, 1.570796, 1.693222],accel_mss,speed_ms,0,blend_radius_m)
  movel([0.125715, -0.674761, -2.795531, -1.242097, 1.570796, 1.696511],accel_mss,speed_ms,0,blend_radius_m)
  movel([0.129133, -0.671312, -2.795926, -1.245151, 1.570796, 1.699929],accel_mss,speed_ms,0,blend_radius_m)
  movel([0.132642, -0.668160, -2.796283, -1.247946, 1.570796, 1.703438],accel_mss,speed_ms,0,blend_radius_m)
  movel([0.136227, -0.665361, -2.796596, -1.250432, 1.570796, 1.707024],accel_mss,speed_ms,0,blend_radius_m)
  movel([0.133977, -0.668260, -2.796272, -1.247858, 1.570796, 1.704773],accel_mss,speed_ms,0,blend_radius_m)
  movel([0.129970, -0.674177, -2.795598, -1.242614, 1.570796, 1.700767],accel_mss,speed_ms,0,blend_radius_m)
  movel([0.128239, -0.677149, -2.795254, -1.239986, 1.570796, 1.699035],accel_mss,speed_ms,0,blend_radius_m)
  movel([0.125396, -0.682957, -2.794570, -1.234862, 1.570796, 1.696193],accel_mss,speed_ms,0,blend_radius_m)
  movel([0.124307, -0.685750, -2.794236, -1.232403, 1.570796, 1.695103],accel_mss,speed_ms,0,blend_radius_m)
  movel([0.123463, -0.688427, -2.793912, -1.230050, 1.570796, 1.694259],accel_mss,speed_ms,0,blend_radius_m)
  speed_ms = 0.005
  movel([0.123463, -0.682196, -2.787256, -1.242937, 1.570796, 1.694259],accel_mss,speed_ms,0,blend_radius_m)
  speed_ms = 0.040
  movel([0.136955, -0.681201, -2.787376, -1.243812, 1.570796, 1.707751],accel_mss,speed_ms,0,blend_radius_m)
  speed_ms = 0.005
  movel([0.136955, -0.687418, -2.794035, -1.230936, 1.570796, 1.707751],accel_mss,speed_ms,0,blend_radius_m)
  speed_ms = 0.025
  movel([0.137370, -0.684148, -2.794428, -1.233813, 1.570796, 1.708167],accel_mss,speed_ms,0,blend_radius_m)
  movel([0.138094, -0.680645, -2.794844, -1.236900, 1.570796, 1.708890],accel_mss,speed_ms,0,blend_radius_m)
  movel([0.139124, -0.676940, -2.795278, -1.240171, 1.570796, 1.709920],accel_mss,speed_ms,0,blend_radius_m)
  movel([0.140459, -0.673070, -2.795725, -1.243593, 1.570796, 1.711255],accel_mss,speed_ms,0,blend_radius_m)
  movel([0.142103, -0.669061, -2.796181, -1.247147, 1.570796, 1.712900],accel_mss,speed_ms,0,blend_radius_m)
  movel([0.144050, -0.664949, -2.796642, -1.250799, 1.570796, 1.714846],accel_mss,speed_ms,0,blend_radius_m)
  movel([0.146296, -0.660763, -2.797103, -1.254523, 1.570796, 1.717093],accel_mss,speed_ms,0,blend_radius_m)
  movel([0.148846, -0.656539, -2.797561, -1.258289, 1.570796, 1.719642],accel_mss,speed_ms,0,blend_radius_m)
  movel([0.157377, -0.643310, -2.798945, -1.270135, 1.570796, 1.728173],accel_mss,speed_ms,0,blend_radius_m)
  movel([0.159091, -0.640259, -2.799253, -1.272876, 1.570796, 1.729888],accel_mss,speed_ms,0,blend_radius_m)
  movel([0.160583, -0.637181, -2.799561, -1.275647, 1.570796, 1.731380],accel_mss,speed_ms,0,blend_radius_m)
  movel([0.161827, -0.634018, -2.799872, -1.278499, 1.570796, 1.732623],accel_mss,speed_ms,0,blend_radius_m)
  movel([0.162797, -0.630693, -2.800196, -1.281500, 1.570796, 1.733593],accel_mss,speed_ms,0,blend_radius_m)
  movel([0.164567, -0.621665, -2.801050, -1.289674, 1.570796, 1.735363],accel_mss,speed_ms,0,blend_radius_m)
  movel([0.165689, -0.617017, -2.801477, -1.293895, 1.570796, 1.736485],accel_mss,speed_ms,0,blend_radius_m)
  movel([0.167508, -0.611983, -2.801929, -1.298477, 1.570796, 1.738304],accel_mss,speed_ms,0,blend_radius_m)
  movel([0.169071, -0.608738, -2.802215, -1.301436, 1.570796, 1.739867],accel_mss,speed_ms,0,blend_radius_m)
  movel([0.170932, -0.605428, -2.802502, -1.304459, 1.570796, 1.741728],accel_mss,speed_ms,0,blend_radius_m)
  movel([0.175378, -0.598683, -2.803074, -1.310632, 1.570796, 1.746174],accel_mss,speed_ms,0,blend_radius_m)
  movel([0.180478, -0.591871, -2.803633, -1.316885, 1.570796, 1.751274],accel_mss,speed_ms,0,blend_radius_m)
  movel([0.185878, -0.585117, -2.804169, -1.323104, 1.570796, 1.756674],accel_mss,speed_ms,0,blend_radius_m)
  movel([0.191243, -0.578632, -2.804666, -1.329091, 1.570796, 1.762039],accel_mss,speed_ms,0,blend_radius_m)
  movel([0.196884, -0.572336, -2.805133, -1.334919, 1.570796, 1.767680],accel_mss,speed_ms,0,blend_radius_m)
  movel([0.199764, -0.569437, -2.805343, -1.337608, 1.570796, 1.770560],accel_mss,speed_ms,0,blend_radius_m)
  movel([0.202667, -0.566788, -2.805532, -1.340068, 1.570796, 1.773464],accel_mss,speed_ms,0,blend_radius_m)
  movel([0.205558, -0.564480, -2.805695, -1.342214, 1.570796, 1.776354],accel_mss,speed_ms,0,blend_radius_m)
  movel([0.208436, -0.562564, -2.805828, -1.343997, 1.570796, 1.779232],accel_mss,speed_ms,0,blend_radius_m)
  speed_ms = 0.005
  movel([0.208436, -0.558258, -2.798950, -1.355181, 1.570796, 1.779232],accel_mss,speed_ms,0,blend_radius_m)
  speed_ms = 0.040
  movel([0.211802, -0.558923, -2.798904, -1.354563, 1.570796, 1.782598],accel_mss,speed_ms,0,blend_radius_m)
  speed_ms = 0.005
  movel([0.211802, -0.563239, -2.805781, -1.343368, 1.570796, 1.782598],accel_mss,speed_ms,0,blend_radius_m)
  speed_ms = 0.025
  movel([0.212871, -0.563332, -2.805775, -1.343283, 1.570796, 1.783668],accel_mss,speed_ms,0,blend_radius_m)
  movel([0.214292, -0.563726, -2.805747, -1.342916, 1.570796, 1.785089],accel_mss,speed_ms,0,blend_radius_m)
  movel([0.216393, -0.565982, -2.805589, -1.340818, 1.570796, 1.787189],accel_mss,speed_ms,0,blend_radius_m)
  movel([0.217015, -0.567593, -2.805475, -1.339321, 1.570796, 1.787812],accel_mss,speed_ms,0,blend_radius_m)
  movel([0.216964, -0.568643, -2.805400, -1.338345, 1.570796, 1.787760],accel_mss,speed_ms,0,blend_radius_m)
  movel([0.216668, -0.569029, -2.805373, -1.337988, 1.570796, 1.787464],accel_mss,speed_ms,0,blend_radius_m)
  movel([0.216115, -0.569251, -2.805357, -1.337782, 1.570796, 1.786911],accel_mss,speed_ms,0,blend_radius_m)
  movel([0.210651, -0.569930, -2.805308, -1.337151, 1.570796, 1.781448],accel_mss,speed_ms,0,blend_radius_m)
  movel([0.207568, -0.570903, -2.805238, -1.336248, 1.570796, 1.778364],accel_mss,speed_ms,0,blend_radius_m)
  movel([0.205881, -0.571788, -2.805173, -1.335427, 1.570796, 1.776678],accel_mss,speed_ms,0,blend_radius_m)
  movel([0.204073, -0.573017, -2.805084, -1.334288, 1.570796, 1.774870],accel_mss,speed_ms,0,blend_radius_m)
  movel([0.202009, -0.574788, -2.804953, -1.332647, 1.570796, 1.772806],accel_mss,speed_ms,0,blend_radius_m)
  movel([0.199978, -0.576794, -2.804804, -1.330791, 1.570796, 1.770774],accel_mss,speed_ms,0,blend_radius_m)
  movel([0.195116, -0.582037, -2.804407, -1.325945, 1.570796, 1.765913],accel_mss,speed_ms,0,blend_radius_m)
  movel([0.190412, -0.587591, -2.803975, -1.320823, 1.570796, 1.761208],accel_mss,speed_ms,0,blend_radius_m)
  movel([0.186005, -0.593283, -2.803518, -1.315587, 1.570796, 1.756801],accel_mss,speed_ms,0,blend_radius_m)
  movel([0.182045, -0.598919, -2.803054, -1.310415, 1.570796, 1.752842],accel_mss,speed_ms,0,blend_radius_m)
  movel([0.184790, -0.602068, -2.802789, -1.307532, 1.570796, 1.755587],accel_mss,speed_ms,0,blend_radius_m)
  movel([0.186760, -0.606053, -2.802448, -1.303888, 1.570796, 1.757556],accel_mss,speed_ms,0,blend_radius_m)
  movel([0.184762, -0.606184, -2.802437, -1.303768, 1.570796, 1.755558],accel_mss,speed_ms,0,blend_radius_m)
  movel([0.182451, -0.606886, -2.802376, -1.303127, 1.570796, 1.753248],accel_mss,speed_ms,0,blend_radius_m)
  movel([0.179901, -0.608145, -2.802267, -1.301977, 1.570796, 1.750697],accel_mss,speed_ms,0,blend_radius_m)
  movel([0.177205, -0.609910, -2.802112, -1.300367, 1.570796, 1.748001],accel_mss,speed_ms,0,blend_radius_m)
  movel([0.175944, -0.611109, -2.802006, -1.299274, 1.570796, 1.746740],accel_mss,speed_ms,0,blend_radius_m)
  movel([0.175442, -0.612313, -2.801900, -1.298176, 1.570796, 1.746238],accel_mss,speed_ms,0,blend_radius_m)
  movel([0.172661, -0.624063, -2.800826, -1.287500, 1.570796, 1.743457],accel_mss,speed_ms,0,blend_radius_m)
  movel([0.170790, -0.630274, -2.800236, -1.281879, 1.570796, 1.741586],accel_mss,speed_ms,0,blend_radius_m)
  movel([0.168470, -0.636785, -2.799600, -1.276004, 1.570796, 1.739266],accel_mss,speed_ms,0,blend_radius_m)
  movel([0.165706, -0.643443, -2.798931, -1.270015, 1.570796, 1.736502],accel_mss,speed_ms,0,blend_radius_m)
  movel([0.162490, -0.650114, -2.798242, -1.264033, 1.570796, 1.733287],accel_mss,speed_ms,0,blend_radius_m)
  movel([0.155700, -0.663543, -2.796797, -1.252048, 1.570796, 1.726496],accel_mss,speed_ms,0,blend_radius_m)
  movel([0.152980, -0.669938, -2.796082, -1.246368, 1.570796, 1.723777],accel_mss,speed_ms,0,blend_radius_m)
  movel([0.151091, -0.676033, -2.795384, -1.240972, 1.570796, 1.721887],accel_mss,speed_ms,0,blend_radius_m)
  speed_ms = 0.005
  movel([0.151091, -0.669973, -2.788701, -1.253715, 1.570796, 1.721887],accel_mss,speed_ms,0,blend_radius_m)
  speed_ms = 0.040
  movel([0.177727, -0.649125, -2.791012, -1.272252, 1.570796, 1.748524],accel_mss,speed_ms,0,blend_radius_m)
  speed_ms = 0.005
  movel([0.177727, -0.654884, -2.797738, -1.259767, 1.570796, 1.748524],accel_mss,speed_ms,0,blend_radius_m)
  speed_ms = 0.025
  movel([0.176157, -0.659877, -2.797200, -1.255312, 1.570796, 1.746954],accel_mss,speed_ms,0,blend_radius_m)
  movel([0.173824, -0.665186, -2.796615, -1.250588, 1.570796, 1.744620],accel_mss,speed_ms,0,blend_radius_m)
  movel([0.170818, -0.670625, -2.796004, -1.245760, 1.570796, 1.741615],accel_mss,speed_ms,0,blend_radius_m)
  movel([0.167242, -0.676020, -2.795385, -1.240984, 1.570796, 1.738039],accel_mss,speed_ms,0,blend_radius_m)
  speed_ms = 0.005
  movel([0.167242, -0.669960, -2.788702, -1.253727, 1.570796, 1.738039],accel_mss,speed_ms,0,blend_radius_m)
  speed_ms = 0.040
  movel([0.161545, -0.667451, -2.788990, -1.255948, 1.570796, 1.732342],accel_mss,speed_ms,0,blend_radius_m)
  speed_ms = 0.005
  movel([0.161545, -0.673475, -2.795679, -1.243235, 1.570796, 1.732342],accel_mss,speed_ms,0,blend_radius_m)
  speed_ms = 0.025
  movel([0.144586, -0.706847, -2.791598, -1.213944, 1.570796, 1.715382],accel_mss,speed_ms,0,blend_radius_m)
  movel([0.143801, -0.708865, -2.791335, -1.212189, 1.570796, 1.714597],accel_mss,speed_ms,0,blend_radius_m)
  movel([0.144115, -0.710540, -2.791115, -1.210733, 1.570796, 1.714911],accel_mss,speed_ms,0,blend_radius_m)
  movel([0.144513, -0.712707, -2.790829, -1.208852, 1.570796, 1.715309],accel_mss,speed_ms,0,blend_radius_m)
  movel([0.144261, -0.715387, -2.790472, -1.206529, 1.570796, 1.715057],accel_mss,speed_ms,0,blend_radius_m)
  speed_ms = 0.005
  movel([0.144261, -0.708800, -2.783877, -1.219711, 1.570796, 1.715057],accel_mss,speed_ms,0,blend_radius_m)
  speed_ms = 0.040
  movel([0.173814, -0.681509, -2.787339, -1.243541, 1.570796, 1.744611],accel_mss,speed_ms,0,blend_radius_m)
  speed_ms = 0.005
  movel([0.173814, -0.687730, -2.793997, -1.230662, 1.570796, 1.744611],accel_mss,speed_ms,0,blend_radius_m)
  speed_ms = 0.025
  movel([0.174212, -0.684772, -2.794353, -1.233264, 1.570796, 1.745008],accel_mss,speed_ms,0,blend_radius_m)
  movel([0.175013, -0.681552, -2.794737, -1.236100, 1.570796, 1.745809],accel_mss,speed_ms,0,blend_radius_m)
  movel([0.176201, -0.678127, -2.795140, -1.239122, 1.570796, 1.746998],accel_mss,speed_ms,0,blend_radius_m)
  movel([0.177775, -0.674535, -2.795557, -1.242297, 1.570796, 1.748571],accel_mss,speed_ms,0,blend_radius_m)
  movel([0.179097, -0.671978, -2.795850, -1.244561, 1.570796, 1.749893],accel_mss,speed_ms,0,blend_radius_m)
  movel([0.180645, -0.669388, -2.796144, -1.246857, 1.570796, 1.751441],accel_mss,speed_ms,0,blend_radius_m)
  movel([0.182421, -0.666862, -2.796428, -1.249099, 1.570796, 1.753217],accel_mss,speed_ms,0,blend_radius_m)
  movel([0.184447, -0.664466, -2.796695, -1.251228, 1.570796, 1.755243],accel_mss,speed_ms,0,blend_radius_m)
  movel([0.186290, -0.662729, -2.796887, -1.252773, 1.570796, 1.757086],accel_mss,speed_ms,0,blend_radius_m)
  movel([0.188308, -0.661220, -2.797053, -1.254116, 1.570796, 1.759104],accel_mss,speed_ms,0,blend_radius_m)
  movel([0.190431, -0.659922, -2.797195, -1.255273, 1.570796, 1.761227],accel_mss,speed_ms,0,blend_radius_m)
  movel([0.192606, -0.658808, -2.797316, -1.256265, 1.570796, 1.763403],accel_mss,speed_ms,0,blend_radius_m)
  movel([0.196844, -0.657041, -2.797507, -1.257841, 1.570796, 1.767641],accel_mss,speed_ms,0,blend_radius_m)
  movel([0.200526, -0.655740, -2.797646, -1.259003, 1.570796, 1.771322],accel_mss,speed_ms,0,blend_radius_m)
  movel([0.197942, -0.656867, -2.797525, -1.257996, 1.570796, 1.768738],accel_mss,speed_ms,0,blend_radius_m)
  movel([0.195252, -0.658503, -2.797349, -1.256537, 1.570796, 1.766048],accel_mss,speed_ms,0,blend_radius_m)
  movel([0.192513, -0.660671, -2.797113, -1.254605, 1.570796, 1.763309],accel_mss,speed_ms,0,blend_radius_m)
  movel([0.189774, -0.663406, -2.796813, -1.252171, 1.570796, 1.760570],accel_mss,speed_ms,0,blend_radius_m)
  movel([0.187593, -0.666090, -2.796515, -1.249784, 1.570796, 1.758390],accel_mss,speed_ms,0,blend_radius_m)
  movel([0.185660, -0.668893, -2.796200, -1.247296, 1.570796, 1.756456],accel_mss,speed_ms,0,blend_radius_m)
  movel([0.184026, -0.671590, -2.795894, -1.244905, 1.570796, 1.754822],accel_mss,speed_ms,0,blend_radius_m)
  movel([0.182637, -0.674251, -2.795590, -1.242549, 1.570796, 1.753433],accel_mss,speed_ms,0,blend_radius_m)
  movel([0.180546, -0.679399, -2.794991, -1.237999, 1.570796, 1.751343],accel_mss,speed_ms,0,blend_radius_m)
  movel([0.179303, -0.684180, -2.794424, -1.233785, 1.570796, 1.750099],accel_mss,speed_ms,0,blend_radius_m)
  movel([0.178810, -0.688798, -2.793867, -1.229723, 1.570796, 1.749606],accel_mss,speed_ms,0,blend_radius_m)
  speed_ms = 0.005
  movel([0.178810, -0.682562, -2.787212, -1.242615, 1.570796, 1.749606],accel_mss,speed_ms,0,blend_radius_m)
  speed_ms = 0.040
  movel([0.186542, -0.669647, -2.788738, -1.254004, 1.570796, 1.757338],accel_mss,speed_ms,0,blend_radius_m)
  speed_ms = 0.005
  movel([0.186542, -0.675702, -2.795422, -1.241265, 1.570796, 1.757338],accel_mss,speed_ms,0,blend_radius_m)
  speed_ms = 0.025
  movel([0.186123, -0.676529, -2.795326, -1.240534, 1.570796, 1.756919],accel_mss,speed_ms,0,blend_radius_m)
  movel([0.185352, -0.677148, -2.795254, -1.239987, 1.570796, 1.756148],accel_mss,speed_ms,0,blend_radius_m)
  movel([0.184878, -0.677034, -2.795267, -1.240088, 1.570796, 1.755674],accel_mss,speed_ms,0,blend_radius_m)
  movel([0.184827, -0.676409, -2.795340, -1.240640, 1.570796, 1.755623],accel_mss,speed_ms,0,blend_radius_m)
  movel([0.185693, -0.674630, -2.795546, -1.242213, 1.570796, 1.756489],accel_mss,speed_ms,0,blend_radius_m)
  movel([0.186300, -0.673835, -2.795637, -1.242917, 1.570796, 1.757097],accel_mss,speed_ms,0,blend_radius_m)
  movel([0.186997, -0.673465, -2.795680, -1.243244, 1.570796, 1.757793],accel_mss,speed_ms,0,blend_radius_m)
  movel([0.187364, -0.673746, -2.795648, -1.242995, 1.570796, 1.758160],accel_mss,speed_ms,0,blend_radius_m)
  movel([0.187006, -0.675276, -2.795471, -1.241641, 1.570796, 1.757803],accel_mss,speed_ms,0,blend_radius_m)
  speed_ms = 0.005
  movel([0.187006, -0.669227, -2.788787, -1.254375, 1.570796, 1.757803],accel_mss,speed_ms,0,blend_radius_m)
  speed_ms = 0.040
  movel([0.185812, -0.687078, -2.786660, -1.238650, 1.570796, 1.756608],accel_mss,speed_ms,0,blend_radius_m)
  speed_ms = 0.005
  movel([0.185812, -0.693376, -2.793306, -1.225707, 1.570796, 1.756608],accel_mss,speed_ms,0,blend_radius_m)
  speed_ms = 0.025
  movel([0.188337, -0.689905, -2.793732, -1.228751, 1.570796, 1.759134],accel_mss,speed_ms,0,blend_radius_m)
  movel([0.190449, -0.686468, -2.794150, -1.231771, 1.570796, 1.761245],accel_mss,speed_ms,0,blend_radius_m)
  movel([0.194703, -0.679523, -2.794976, -1.237890, 1.570796, 1.765499],accel_mss,speed_ms,0,blend_radius_m)
  movel([0.198340, -0.674643, -2.795544, -1.242202, 1.570796, 1.769136],accel_mss,speed_ms,0,blend_radius_m)
  movel([0.210611, -0.659906, -2.797196, -1.255287, 1.570796, 1.781407],accel_mss,speed_ms,0,blend_radius_m)
  movel([0.212945, -0.656707, -2.797543, -1.258139, 1.570796, 1.783741],accel_mss,speed_ms,0,blend_radius_m)
  movel([0.213697, -0.655215, -2.797703, -1.259472, 1.570796, 1.784493],accel_mss,speed_ms,0,blend_radius_m)
  movel([0.213863, -0.654040, -2.797828, -1.260521, 1.570796, 1.784659],accel_mss,speed_ms,0,blend_radius_m)
  movel([0.213139, -0.653417, -2.797894, -1.261078, 1.570796, 1.783936],accel_mss,speed_ms,0,blend_radius_m)
  movel([0.211867, -0.653497, -2.797886, -1.261007, 1.570796, 1.782663],accel_mss,speed_ms,0,blend_radius_m)
  movel([0.209782, -0.654027, -2.797829, -1.260533, 1.570796, 1.780579],accel_mss,speed_ms,0,blend_radius_m)
  movel([0.207684, -0.655022, -2.797723, -1.259644, 1.570796, 1.778481],accel_mss,speed_ms,0,blend_radius_m)
  movel([0.205428, -0.656590, -2.797555, -1.258244, 1.570796, 1.776225],accel_mss,speed_ms,0,blend_radius_m)
  movel([0.202879, -0.658830, -2.797313, -1.256246, 1.570796, 1.773676],accel_mss,speed_ms,0,blend_radius_m)
  movel([0.200205, -0.661618, -2.797009, -1.253762, 1.570796, 1.771001],accel_mss,speed_ms,0,blend_radius_m)
  movel([0.197622, -0.664749, -2.796664, -1.250976, 1.570796, 1.768418],accel_mss,speed_ms,0,blend_radius_m)
  movel([0.195151, -0.668111, -2.796288, -1.247990, 1.570796, 1.765947],accel_mss,speed_ms,0,blend_radius_m)
  movel([0.192804, -0.671617, -2.795891, -1.244881, 1.570796, 1.763600],accel_mss,speed_ms,0,blend_radius_m)
  movel([0.188561, -0.678624, -2.795082, -1.238683, 1.570796, 1.759357],accel_mss,speed_ms,0,blend_radius_m)
  movel([0.185008, -0.684987, -2.794328, -1.233074, 1.570796, 1.755804],accel_mss,speed_ms,0,blend_radius_m)
  movel([0.178825, -0.696641, -2.792899, -1.222848, 1.570796, 1.749621],accel_mss,speed_ms,0,blend_radius_m)
  movel([0.176582, -0.700497, -2.792413, -1.219479, 1.570796, 1.747378],accel_mss,speed_ms,0,blend_radius_m)
  movel([0.174060, -0.704353, -2.791921, -1.216116, 1.570796, 1.744857],accel_mss,speed_ms,0,blend_radius_m)
  movel([0.171242, -0.708085, -2.791437, -1.212867, 1.570796, 1.742038],accel_mss,speed_ms,0,blend_radius_m)
  movel([0.168189, -0.711499, -2.790989, -1.209900, 1.570796, 1.738986],accel_mss,speed_ms,0,blend_radius_m)
  movel([0.164961, -0.714407, -2.790603, -1.207379, 1.570796, 1.735757],accel_mss,speed_ms,0,blend_radius_m)
  movel([0.167425, -0.713090, -2.790779, -1.208521, 1.570796, 1.738222],accel_mss,speed_ms,0,blend_radius_m)
  movel([0.169955, -0.711497, -2.790989, -1.209902, 1.570796, 1.740751],accel_mss,speed_ms,0,blend_radius_m)
  movel([0.172526, -0.709637, -2.791234, -1.211518, 1.570796, 1.743323],accel_mss,speed_ms,0,blend_radius_m)
  movel([0.175099, -0.707544, -2.791508, -1.213338, 1.570796, 1.745895],accel_mss,speed_ms,0,blend_radius_m)
  movel([0.174856, -0.710252, -2.791153, -1.210984, 1.570796, 1.745652],accel_mss,speed_ms,0,blend_radius_m)
  movel([0.174158, -0.713247, -2.790758, -1.208384, 1.570796, 1.744954],accel_mss,speed_ms,0,blend_radius_m)
  movel([0.173033, -0.716449, -2.790330, -1.205610, 1.570796, 1.743829],accel_mss,speed_ms,0,blend_radius_m)
  movel([0.171507, -0.719781, -2.789880, -1.202728, 1.570796, 1.742303],accel_mss,speed_ms,0,blend_radius_m)
  movel([0.174336, -0.716065, -2.790382, -1.205943, 1.570796, 1.745132],accel_mss,speed_ms,0,blend_radius_m)
  movel([0.176844, -0.712276, -2.790886, -1.209226, 1.570796, 1.747641],accel_mss,speed_ms,0,blend_radius_m)
  movel([0.179054, -0.708441, -2.791391, -1.212558, 1.570796, 1.749850],accel_mss,speed_ms,0,blend_radius_m)
  movel([0.180999, -0.704580, -2.791891, -1.215918, 1.570796, 1.751796],accel_mss,speed_ms,0,blend_radius_m)
  movel([0.180935, -0.706340, -2.791664, -1.214385, 1.570796, 1.751731],accel_mss,speed_ms,0,blend_radius_m)
  movel([0.180430, -0.708544, -2.791377, -1.212468, 1.570796, 1.751227],accel_mss,speed_ms,0,blend_radius_m)
  movel([0.176636, -0.719179, -2.789962, -1.203248, 1.570796, 1.747432],accel_mss,speed_ms,0,blend_radius_m)
  movel([0.175905, -0.721669, -2.789623, -1.201097, 1.570796, 1.746701],accel_mss,speed_ms,0,blend_radius_m)
  movel([0.175524, -0.723835, -2.789325, -1.199229, 1.570796, 1.746321],accel_mss,speed_ms,0,blend_radius_m)
  movel([0.177223, -0.720029, -2.789846, -1.202514, 1.570796, 1.748019],accel_mss,speed_ms,0,blend_radius_m)
  movel([0.179115, -0.716392, -2.790338, -1.205660, 1.570796, 1.749911],accel_mss,speed_ms,0,blend_radius_m)
  movel([0.183325, -0.709416, -2.791263, -1.211710, 1.570796, 1.754121],accel_mss,speed_ms,0,blend_radius_m)
  movel([0.187856, -0.702448, -2.792165, -1.217776, 1.570796, 1.758653],accel_mss,speed_ms,0,blend_radius_m)
  movel([0.192430, -0.694998, -2.793105, -1.224287, 1.570796, 1.763227],accel_mss,speed_ms,0,blend_radius_m)
  movel([0.194843, -0.690396, -2.793672, -1.228321, 1.570796, 1.765639],accel_mss,speed_ms,0,blend_radius_m)
  movel([0.196435, -0.687784, -2.793990, -1.230614, 1.570796, 1.767231],accel_mss,speed_ms,0,blend_radius_m)
  movel([0.197216, -0.686784, -2.794111, -1.231494, 1.570796, 1.768012],accel_mss,speed_ms,0,blend_radius_m)
  movel([0.197953, -0.686124, -2.794191, -1.232074, 1.570796, 1.768749],accel_mss,speed_ms,0,blend_radius_m)
  movel([0.198592, -0.685875, -2.794221, -1.232293, 1.570796, 1.769389],accel_mss,speed_ms,0,blend_radius_m)
  movel([0.199114, -0.685981, -2.794208, -1.232200, 1.570796, 1.769910],accel_mss,speed_ms,0,blend_radius_m)
  movel([0.199801, -0.686959, -2.794090, -1.231340, 1.570796, 1.770597],accel_mss,speed_ms,0,blend_radius_m)
  movel([0.199974, -0.688497, -2.793904, -1.229988, 1.570796, 1.770770],accel_mss,speed_ms,0,blend_radius_m)
  movel([0.199596, -0.690038, -2.793716, -1.228635, 1.570796, 1.770392],accel_mss,speed_ms,0,blend_radius_m)
  movel([0.202193, -0.684285, -2.794412, -1.233692, 1.570796, 1.772990],accel_mss,speed_ms,0,blend_radius_m)
  movel([0.204277, -0.678686, -2.795074, -1.238629, 1.570796, 1.775073],accel_mss,speed_ms,0,blend_radius_m)
  movel([0.205821, -0.673326, -2.795696, -1.243367, 1.570796, 1.776618],accel_mss,speed_ms,0,blend_radius_m)
  movel([0.206788, -0.668289, -2.796268, -1.247832, 1.570796, 1.777584],accel_mss,speed_ms,0,blend_radius_m)
  speed_ms = 0.005
  movel([0.206788, -0.662338, -2.789569, -1.260482, 1.570796, 1.777584],accel_mss,speed_ms,0,blend_radius_m)
  speed_ms = 0.040
  movel([0.211773, -0.661776, -2.789632, -1.260981, 1.570796, 1.782569],accel_mss,speed_ms,0,blend_radius_m)
  speed_ms = 0.005
  movel([0.211773, -0.667718, -2.796332, -1.248338, 1.570796, 1.782569],accel_mss,speed_ms,0,blend_radius_m)
  speed_ms = 0.025
  movel([0.214738, -0.667099, -2.796402, -1.248888, 1.570796, 1.785534],accel_mss,speed_ms,0,blend_radius_m)
  movel([0.215823, -0.667358, -2.796373, -1.248658, 1.570796, 1.786620],accel_mss,speed_ms,0,blend_radius_m)
  movel([0.216375, -0.668255, -2.796272, -1.247862, 1.570796, 1.787171],accel_mss,speed_ms,0,blend_radius_m)
  movel([0.216315, -0.669527, -2.796129, -1.246733, 1.570796, 1.787112],accel_mss,speed_ms,0,blend_radius_m)
  movel([0.210190, -0.693695, -2.793266, -1.225428, 1.570796, 1.780986],accel_mss,speed_ms,0,blend_radius_m)
  movel([0.209662, -0.695453, -2.793048, -1.223888, 1.570796, 1.780459],accel_mss,speed_ms,0,blend_radius_m)
  movel([0.208882, -0.697311, -2.792816, -1.222263, 1.570796, 1.779679],accel_mss,speed_ms,0,blend_radius_m)
  movel([0.207798, -0.699066, -2.792595, -1.220728, 1.570796, 1.778594],accel_mss,speed_ms,0,blend_radius_m)
  movel([0.206377, -0.700506, -2.792412, -1.219471, 1.570796, 1.777173],accel_mss,speed_ms,0,blend_radius_m)
  movel([0.205028, -0.701234, -2.792320, -1.218836, 1.570796, 1.775825],accel_mss,speed_ms,0,blend_radius_m)
  movel([0.202542, -0.701871, -2.792239, -1.218280, 1.570796, 1.773338],accel_mss,speed_ms,0,blend_radius_m)
  movel([0.201197, -0.702655, -2.792138, -1.217596, 1.570796, 1.771993],accel_mss,speed_ms,0,blend_radius_m)
  movel([0.199617, -0.704358, -2.791920, -1.216111, 1.570796, 1.770413],accel_mss,speed_ms,0,blend_radius_m)
  movel([0.198216, -0.706321, -2.791666, -1.214402, 1.570796, 1.769012],accel_mss,speed_ms,0,blend_radius_m)
  movel([0.196444, -0.708566, -2.791374, -1.212449, 1.570796, 1.767240],accel_mss,speed_ms,0,blend_radius_m)
  movel([0.194510, -0.710604, -2.791107, -1.210678, 1.570796, 1.765306],accel_mss,speed_ms,0,blend_radius_m)
  movel([0.192490, -0.712386, -2.790872, -1.209131, 1.570796, 1.763286],accel_mss,speed_ms,0,blend_radius_m)
  movel([0.190451, -0.713868, -2.790675, -1.207846, 1.570796, 1.761247],accel_mss,speed_ms,0,blend_radius_m)
  movel([0.188462, -0.715009, -2.790523, -1.206857, 1.570796, 1.759258],accel_mss,speed_ms,0,blend_radius_m)
  movel([0.186605, -0.715752, -2.790424, -1.206214, 1.570796, 1.757401],accel_mss,speed_ms,0,blend_radius_m)
  movel([0.184943, -0.716066, -2.790381, -1.205942, 1.570796, 1.755739],accel_mss,speed_ms,0,blend_radius_m)
  movel([0.183550, -0.715889, -2.790405, -1.206095, 1.570796, 1.754346],accel_mss,speed_ms,0,blend_radius_m)
  speed_ms = 0.005
  movel([0.183550, -0.709295, -2.783811, -1.219282, 1.570796, 1.754346],accel_mss,speed_ms,0,blend_radius_m)
  speed_ms = 0.040
  movel([0.168134, -0.734536, -2.780294, -1.197559, 1.570796, 1.738930],accel_mss,speed_ms,0,blend_radius_m)
  speed_ms = 0.005
  movel([0.168134, -0.741447, -2.786825, -1.184117, 1.570796, 1.738930],accel_mss,speed_ms,0,blend_radius_m)
  speed_ms = 0.025
  movel([0.167046, -0.761688, -2.783765, -1.166936, 1.570796, 1.737842],accel_mss,speed_ms,0,blend_radius_m)
  movel([0.166647, -0.764319, -2.783353, -1.164717, 1.570796, 1.737443],accel_mss,speed_ms,0,blend_radius_m)
  movel([0.166087, -0.765743, -2.783128, -1.163518, 1.570796, 1.736883],accel_mss,speed_ms,0,blend_radius_m)
  movel([0.165160, -0.767172, -2.782901, -1.162316, 1.570796, 1.735956],accel_mss,speed_ms,0,blend_radius_m)
  movel([0.162600, -0.769984, -2.782452, -1.159953, 1.570796, 1.733397],accel_mss,speed_ms,0,blend_radius_m)
  movel([0.161837, -0.771545, -2.782201, -1.158643, 1.570796, 1.732633],accel_mss,speed_ms,0,blend_radius_m)
  movel([0.161582, -0.772959, -2.781973, -1.157457, 1.570796, 1.732378],accel_mss,speed_ms,0,blend_radius_m)
  movel([0.161838, -0.774858, -2.781665, -1.155866, 1.570796, 1.732634],accel_mss,speed_ms,0,blend_radius_m)
  movel([0.162673, -0.776315, -2.781427, -1.154647, 1.570796, 1.733469],accel_mss,speed_ms,0,blend_radius_m)
  movel([0.164736, -0.778724, -2.781031, -1.152634, 1.570796, 1.735533],accel_mss,speed_ms,0,blend_radius_m)
  movel([0.165611, -0.780807, -2.780687, -1.150895, 1.570796, 1.736407],accel_mss,speed_ms,0,blend_radius_m)
  movel([0.166290, -0.784250, -2.780113, -1.148026, 1.570796, 1.737087],accel_mss,speed_ms,0,blend_radius_m)
  movel([0.166249, -0.786044, -2.779811, -1.146534, 1.570796, 1.737046],accel_mss,speed_ms,0,blend_radius_m)
  movel([0.165788, -0.787668, -2.779536, -1.145184, 1.570796, 1.736584],accel_mss,speed_ms,0,blend_radius_m)
  movel([0.165360, -0.788357, -2.779420, -1.144613, 1.570796, 1.736156],accel_mss,speed_ms,0,blend_radius_m)
  movel([0.164784, -0.788940, -2.779321, -1.144128, 1.570796, 1.735580],accel_mss,speed_ms,0,blend_radius_m)
  movel([0.164041, -0.789396, -2.779243, -1.143750, 1.570796, 1.734838],accel_mss,speed_ms,0,blend_radius_m)
  movel([0.163120, -0.789698, -2.779191, -1.143500, 1.570796, 1.733916],accel_mss,speed_ms,0,blend_radius_m)
  movel([0.162810, -0.791365, -2.778907, -1.142118, 1.570796, 1.733606],accel_mss,speed_ms,0,blend_radius_m)
  movel([0.162912, -0.792992, -2.778627, -1.140770, 1.570796, 1.733708],accel_mss,speed_ms,0,blend_radius_m)
  movel([0.163975, -0.796040, -2.778100, -1.138250, 1.570796, 1.734772],accel_mss,speed_ms,0,blend_radius_m)
  movel([0.165590, -0.798624, -2.777649, -1.136116, 1.570796, 1.736386],accel_mss,speed_ms,0,blend_radius_m)
  movel([0.167059, -0.800512, -2.777317, -1.134560, 1.570796, 1.737855],accel_mss,speed_ms,0,blend_radius_m)
  movel([0.169114, -0.802149, -2.777028, -1.133212, 1.570796, 1.739910],accel_mss,speed_ms,0,blend_radius_m)
  movel([0.171552, -0.803508, -2.776787, -1.132095, 1.570796, 1.742348],accel_mss,speed_ms,0,blend_radius_m)
  movel([0.173567, -0.805283, -2.776470, -1.130636, 1.570796, 1.744364],accel_mss,speed_ms,0,blend_radius_m)
  movel([0.174168, -0.806534, -2.776246, -1.129609, 1.570796, 1.744964],accel_mss,speed_ms,0,blend_radius_m)
  movel([0.174361, -0.808144, -2.775956, -1.128289, 1.570796, 1.745157],accel_mss,speed_ms,0,blend_radius_m)
  movel([0.174197, -0.809153, -2.775774, -1.127462, 1.570796, 1.744993],accel_mss,speed_ms,0,blend_radius_m)
  movel([0.173762, -0.810281, -2.775570, -1.126538, 1.570796, 1.744559],accel_mss,speed_ms,0,blend_radius_m)
  movel([0.173098, -0.811298, -2.775385, -1.125706, 1.570796, 1.743895],accel_mss,speed_ms,0,blend_radius_m)
  movel([0.172238, -0.811991, -2.775259, -1.125139, 1.570796, 1.743034],accel_mss,speed_ms,0,blend_radius_m)
  movel([0.171591, -0.812126, -2.775234, -1.125029, 1.570796, 1.742387],accel_mss,speed_ms,0,blend_radius_m)
  movel([0.171082, -0.811992, -2.775259, -1.125139, 1.570796, 1.741878],accel_mss,speed_ms,0,blend_radius_m)
  movel([0.166878, -0.809773, -2.775662, -1.126954, 1.570796, 1.737674],accel_mss,speed_ms,0,blend_radius_m)
  movel([0.165032, -0.808331, -2.775923, -1.128135, 1.570796, 1.735828],accel_mss,speed_ms,0,blend_radius_m)
  movel([0.163371, -0.806664, -2.776223, -1.129502, 1.570796, 1.734167],accel_mss,speed_ms,0,blend_radius_m)
  movel([0.162682, -0.807839, -2.776011, -1.128539, 1.570796, 1.733478],accel_mss,speed_ms,0,blend_radius_m)
  movel([0.162225, -0.808983, -2.775805, -1.127601, 1.570796, 1.733021],accel_mss,speed_ms,0,blend_radius_m)
  movel([0.161921, -0.811165, -2.775409, -1.125815, 1.570796, 1.732718],accel_mss,speed_ms,0,blend_radius_m)
  movel([0.162270, -0.813189, -2.775040, -1.124160, 1.570796, 1.733067],accel_mss,speed_ms,0,blend_radius_m)
  movel([0.163102, -0.815028, -2.774702, -1.122659, 1.570796, 1.733899],accel_mss,speed_ms,0,blend_radius_m)
  movel([0.165470, -0.818094, -2.774135, -1.120160, 1.570796, 1.736266],accel_mss,speed_ms,0,blend_radius_m)
  movel([0.167615, -0.820163, -2.773750, -1.118476, 1.570796, 1.738411],accel_mss,speed_ms,0,blend_radius_m)
  movel([0.168264, -0.821085, -2.773577, -1.117726, 1.570796, 1.739061],accel_mss,speed_ms,0,blend_radius_m)
  movel([0.168336, -0.821736, -2.773455, -1.117197, 1.570796, 1.739132],accel_mss,speed_ms,0,blend_radius_m)
  movel([0.168092, -0.822568, -2.773299, -1.116522, 1.570796, 1.738888],accel_mss,speed_ms,0,blend_radius_m)
  movel([0.167525, -0.823509, -2.773122, -1.115759, 1.570796, 1.738321],accel_mss,speed_ms,0,blend_radius_m)
  movel([0.166905, -0.824128, -2.773005, -1.115256, 1.570796, 1.737702],accel_mss,speed_ms,0,blend_radius_m)
  movel([0.165611, -0.824721, -2.772893, -1.114776, 1.570796, 1.736408],accel_mss,speed_ms,0,blend_radius_m)
  movel([0.163841, -0.825331, -2.772777, -1.114281, 1.570796, 1.734637],accel_mss,speed_ms,0,blend_radius_m)
  movel([0.163392, -0.825806, -2.772687, -1.113896, 1.570796, 1.734188],accel_mss,speed_ms,0,blend_radius_m)
  movel([0.163003, -0.826613, -2.772533, -1.113243, 1.570796, 1.733800],accel_mss,speed_ms,0,blend_radius_m)
  movel([0.162866, -0.827422, -2.772379, -1.112588, 1.570796, 1.733662],accel_mss,speed_ms,0,blend_radius_m)
  movel([0.163142, -0.828968, -2.772083, -1.111338, 1.570796, 1.733938],accel_mss,speed_ms,0,blend_radius_m)
  movel([0.164334, -0.831288, -2.771637, -1.109464, 1.570796, 1.735130],accel_mss,speed_ms,0,blend_radius_m)
  movel([0.167273, -0.835790, -2.770762, -1.105837, 1.570796, 1.738069],accel_mss,speed_ms,0,blend_radius_m)
  movel([0.170319, -0.840155, -2.769903, -1.102331, 1.570796, 1.741115],accel_mss,speed_ms,0,blend_radius_m)
  movel([0.170739, -0.841223, -2.769691, -1.101474, 1.570796, 1.741535],accel_mss,speed_ms,0,blend_radius_m)
  movel([0.170851, -0.842548, -2.769427, -1.100414, 1.570796, 1.741647],accel_mss,speed_ms,0,blend_radius_m)
  movel([0.170481, -0.844023, -2.769133, -1.099233, 1.570796, 1.741277],accel_mss,speed_ms,0,blend_radius_m)
  movel([0.170070, -0.844777, -2.768981, -1.098630, 1.570796, 1.740866],accel_mss,speed_ms,0,blend_radius_m)
  movel([0.168821, -0.846128, -2.768710, -1.097551, 1.570796, 1.739618],accel_mss,speed_ms,0,blend_radius_m)
  movel([0.168185, -0.846534, -2.768628, -1.097227, 1.570796, 1.738981],accel_mss,speed_ms,0,blend_radius_m)
  movel([0.166974, -0.846862, -2.768562, -1.096965, 1.570796, 1.737771],accel_mss,speed_ms,0,blend_radius_m)
  movel([0.165901, -0.846708, -2.768593, -1.097088, 1.570796, 1.736697],accel_mss,speed_ms,0,blend_radius_m)
  movel([0.165025, -0.846252, -2.768685, -1.097452, 1.570796, 1.735821],accel_mss,speed_ms,0,blend_radius_m)
  movel([0.160516, -0.842741, -2.769389, -1.100259, 1.570796, 1.731312],accel_mss,speed_ms,0,blend_radius_m)
  movel([0.156319, -0.838830, -2.770165, -1.103394, 1.570796, 1.727115],accel_mss,speed_ms,0,blend_radius_m)
  movel([0.152457, -0.834511, -2.771012, -1.106867, 1.570796, 1.723253],accel_mss,speed_ms,0,blend_radius_m)
  movel([0.148937, -0.829784, -2.771926, -1.110678, 1.570796, 1.719734],accel_mss,speed_ms,0,blend_radius_m)
  movel([0.147785, -0.827869, -2.772294, -1.112227, 1.570796, 1.718581],accel_mss,speed_ms,0,blend_radius_m)
  movel([0.147080, -0.825537, -2.772738, -1.114114, 1.570796, 1.717877],accel_mss,speed_ms,0,blend_radius_m)
  movel([0.147019, -0.823867, -2.773054, -1.115468, 1.570796, 1.717815],accel_mss,speed_ms,0,blend_radius_m)
  movel([0.147185, -0.822037, -2.773399, -1.116953, 1.570796, 1.717981],accel_mss,speed_ms,0,blend_radius_m)
  movel([0.147900, -0.818122, -2.774130, -1.120137, 1.570796, 1.718696],accel_mss,speed_ms,0,blend_radius_m)
  movel([0.151798, -0.803301, -2.776823, -1.132265, 1.570796, 1.722594],accel_mss,speed_ms,0,blend_radius_m)
  movel([0.152566, -0.799255, -2.777538, -1.135596, 1.570796, 1.723363],accel_mss,speed_ms,0,blend_radius_m)
  movel([0.152817, -0.795838, -2.778135, -1.138416, 1.570796, 1.723614],accel_mss,speed_ms,0,blend_radius_m)
  movel([0.152686, -0.794485, -2.778369, -1.139535, 1.570796, 1.723483],accel_mss,speed_ms,0,blend_radius_m)
  movel([0.152339, -0.793440, -2.778550, -1.140399, 1.570796, 1.723136],accel_mss,speed_ms,0,blend_radius_m)
  movel([0.151757, -0.792746, -2.778669, -1.140974, 1.570796, 1.722554],accel_mss,speed_ms,0,blend_radius_m)
  movel([0.150915, -0.792452, -2.778720, -1.141217, 1.570796, 1.721711],accel_mss,speed_ms,0,blend_radius_m)
  movel([0.149073, -0.792590, -2.778696, -1.141103, 1.570796, 1.719869],accel_mss,speed_ms,0,blend_radius_m)
  movel([0.148262, -0.792524, -2.778708, -1.141157, 1.570796, 1.719058],accel_mss,speed_ms,0,blend_radius_m)
  movel([0.147749, -0.792074, -2.778785, -1.141530, 1.570796, 1.718546],accel_mss,speed_ms,0,blend_radius_m)
  movel([0.147797, -0.790649, -2.779029, -1.142711, 1.570796, 1.718594],accel_mss,speed_ms,0,blend_radius_m)
  movel([0.148457, -0.788834, -2.779339, -1.144216, 1.570796, 1.719253],accel_mss,speed_ms,0,blend_radius_m)
  movel([0.150783, -0.782939, -2.780332, -1.149118, 1.570796, 1.721580],accel_mss,speed_ms,0,blend_radius_m)
  movel([0.152808, -0.777156, -2.781289, -1.153943, 1.570796, 1.723604],accel_mss,speed_ms,0,blend_radius_m)
  movel([0.154569, -0.771459, -2.782215, -1.158715, 1.570796, 1.725366],accel_mss,speed_ms,0,blend_radius_m)
  movel([0.156106, -0.765829, -2.783114, -1.163446, 1.570796, 1.726902],accel_mss,speed_ms,0,blend_radius_m)
  movel([0.158705, -0.754677, -2.784848, -1.172864, 1.570796, 1.729502],accel_mss,speed_ms,0,blend_radius_m)
  movel([0.160963, -0.743502, -2.786523, -1.182364, 1.570796, 1.731759],accel_mss,speed_ms,0,blend_radius_m)
  speed_ms = 0.005
  movel([0.160963, -0.736566, -2.779998, -1.195825, 1.570796, 1.731759],accel_mss,speed_ms,0,blend_radius_m)
  speed_ms = 0.040
  movel([0.150594, -0.766063, -2.775464, -1.170862, 1.570796, 1.721391],accel_mss,speed_ms,0,blend_radius_m)
  speed_ms = 0.005
  movel([0.150594, -0.773341, -2.781911, -1.157137, 1.570796, 1.721391],accel_mss,speed_ms,0,blend_radius_m)
  speed_ms = 0.025
  movel([0.144726, -0.781708, -2.780537, -1.150144, 1.570796, 1.715522],accel_mss,speed_ms,0,blend_radius_m)
  movel([0.138704, -0.789881, -2.779160, -1.143348, 1.570796, 1.709501],accel_mss,speed_ms,0,blend_radius_m)
  movel([0.132543, -0.797853, -2.777783, -1.136752, 1.570796, 1.703339],accel_mss,speed_ms,0,blend_radius_m)
  movel([0.126261, -0.805599, -2.776414, -1.130377, 1.570796, 1.697058],accel_mss,speed_ms,0,blend_radius_m)
  movel([0.130947, -0.797897, -2.777776, -1.136716, 1.570796, 1.701744],accel_mss,speed_ms,0,blend_radius_m)
  movel([0.135271, -0.790094, -2.779124, -1.143171, 1.570796, 1.706068],accel_mss,speed_ms,0,blend_radius_m)
  movel([0.139199, -0.782245, -2.780448, -1.149696, 1.570796, 1.709995],accel_mss,speed_ms,0,blend_radius_m)
  movel([0.142697, -0.774406, -2.781738, -1.156244, 1.570796, 1.713493],accel_mss,speed_ms,0,blend_radius_m)
  movel([0.137758, -0.781285, -2.780608, -1.150496, 1.570796, 1.708554],accel_mss,speed_ms,0,blend_radius_m)
  movel([0.132705, -0.788015, -2.779478, -1.144896, 1.570796, 1.703501],accel_mss,speed_ms,0,blend_radius_m)
  movel([0.127537, -0.794596, -2.778350, -1.139443, 1.570796, 1.698334],accel_mss,speed_ms,0,blend_radius_m)
  movel([0.122271, -0.801005, -2.777230, -1.134154, 1.570796, 1.693068],accel_mss,speed_ms,0,blend_radius_m)
  movel([0.116374, -0.807995, -2.775983, -1.128411, 1.570796, 1.687170],accel_mss,speed_ms,0,blend_radius_m)
  movel([0.110781, -0.815080, -2.774693, -1.122616, 1.570796, 1.681577],accel_mss,speed_ms,0,blend_radius_m)
  movel([0.108244, -0.818744, -2.774014, -1.119630, 1.570796, 1.679040],accel_mss,speed_ms,0,blend_radius_m)
  movel([0.106002, -0.822453, -2.773321, -1.116616, 1.570796, 1.676798],accel_mss,speed_ms,0,blend_radius_m)
  movel([0.104188, -0.826109, -2.772629, -1.113651, 1.570796, 1.674985],accel_mss,speed_ms,0,blend_radius_m)
  movel([0.102912, -0.829621, -2.771958, -1.110810, 1.570796, 1.673708],accel_mss,speed_ms,0,blend_radius_m)
  movel([0.103673, -0.825626, -2.772721, -1.114042, 1.570796, 1.674469],accel_mss,speed_ms,0,blend_radius_m)
  movel([0.104773, -0.821357, -2.773526, -1.117505, 1.570796, 1.675570],accel_mss,speed_ms,0,blend_radius_m)
  movel([0.106194, -0.816871, -2.774362, -1.121156, 1.570796, 1.676990],accel_mss,speed_ms,0,blend_radius_m)
  movel([0.107911, -0.812220, -2.775217, -1.124952, 1.570796, 1.678707],accel_mss,speed_ms,0,blend_radius_m)
  movel([0.109899, -0.807466, -2.776078, -1.128844, 1.570796, 1.680696],accel_mss,speed_ms,0,blend_radius_m)
  movel([0.112139, -0.802663, -2.776937, -1.132790, 1.570796, 1.682936],accel_mss,speed_ms,0,blend_radius_m)
  movel([0.114604, -0.797873, -2.777780, -1.136736, 1.570796, 1.685401],accel_mss,speed_ms,0,blend_radius_m)
  movel([0.117266, -0.793163, -2.778597, -1.140628, 1.570796, 1.688063],accel_mss,speed_ms,0,blend_radius_m)
  movel([0.112338, -0.800639, -2.777294, -1.134455, 1.570796, 1.683134],accel_mss,speed_ms,0,blend_radius_m)
  movel([0.107760, -0.808080, -2.775968, -1.128341, 1.570796, 1.678556],accel_mss,speed_ms,0,blend_radius_m)
  movel([0.103507, -0.815470, -2.774621, -1.122298, 1.570796, 1.674303],accel_mss,speed_ms,0,blend_radius_m)
  movel([0.099554, -0.822791, -2.773257, -1.116341, 1.570796, 1.670351],accel_mss,speed_ms,0,blend_radius_m)
  movel([0.095883, -0.830023, -2.771881, -1.110486, 1.570796, 1.666679],accel_mss,speed_ms,0,blend_radius_m)
  movel([0.092464, -0.837152, -2.770495, -1.104742, 1.570796, 1.663260],accel_mss,speed_ms,0,blend_radius_m)
  movel([0.086284, -0.851039, -2.767713, -1.093636, 1.570796, 1.657080],accel_mss,speed_ms,0,blend_radius_m)
  movel([0.087878, -0.846408, -2.768653, -1.097328, 1.570796, 1.658675],accel_mss,speed_ms,0,blend_radius_m)
  movel([0.089011, -0.841628, -2.769611, -1.101150, 1.570796, 1.659807],accel_mss,speed_ms,0,blend_radius_m)
  movel([0.090902, -0.832403, -2.771421, -1.108565, 1.570796, 1.661699],accel_mss,speed_ms,0,blend_radius_m)
  movel([0.092098, -0.828155, -2.772239, -1.111995, 1.570796, 1.662894],accel_mss,speed_ms,0,blend_radius_m)
  movel([0.093464, -0.824221, -2.772987, -1.115181, 1.570796, 1.664260],accel_mss,speed_ms,0,blend_radius_m)
  movel([0.096953, -0.815868, -2.774547, -1.121973, 1.570796, 1.667749],accel_mss,speed_ms,0,blend_radius_m)
  movel([0.096140, -0.817128, -2.774315, -1.120946, 1.570796, 1.666936],accel_mss,speed_ms,0,blend_radius_m)
  movel([0.094705, -0.818823, -2.774000, -1.119566, 1.570796, 1.665501],accel_mss,speed_ms,0,blend_radius_m)
  movel([0.086526, -0.827146, -2.772432, -1.112811, 1.570796, 1.657322],accel_mss,speed_ms,0,blend_radius_m)
  movel([0.083608, -0.830282, -2.771831, -1.110276, 1.570796, 1.654405],accel_mss,speed_ms,0,blend_radius_m)
  movel([0.080476, -0.834575, -2.770999, -1.106814, 1.570796, 1.651272],accel_mss,speed_ms,0,blend_radius_m)
  movel([0.077643, -0.839061, -2.770119, -1.103209, 1.570796, 1.648440],accel_mss,speed_ms,0,blend_radius_m)
  movel([0.072660, -0.847991, -2.768333, -1.096064, 1.570796, 1.643456],accel_mss,speed_ms,0,blend_radius_m)
  movel([0.074474, -0.843464, -2.769244, -1.099680, 1.570796, 1.645271],accel_mss,speed_ms,0,blend_radius_m)
  movel([0.075968, -0.838998, -2.770132, -1.103259, 1.570796, 1.646764],accel_mss,speed_ms,0,blend_radius_m)
  movel([0.078867, -0.830022, -2.771881, -1.110486, 1.570796, 1.649663],accel_mss,speed_ms,0,blend_radius_m)
  movel([0.080779, -0.825214, -2.772799, -1.114376, 1.570796, 1.651575],accel_mss,speed_ms,0,blend_radius_m)
  movel([0.083046, -0.820267, -2.773731, -1.118391, 1.570796, 1.653842],accel_mss,speed_ms,0,blend_radius_m)
  movel([0.088389, -0.810043, -2.775613, -1.126733, 1.570796, 1.659185],accel_mss,speed_ms,0,blend_radius_m)
  movel([0.100262, -0.789274, -2.779264, -1.143851, 1.570796, 1.671058],accel_mss,speed_ms,0,blend_radius_m)
  movel([0.095207, -0.793865, -2.778476, -1.140048, 1.570796, 1.666004],accel_mss,speed_ms,0,blend_radius_m)
  movel([0.090287, -0.798705, -2.777634, -1.136049, 1.570796, 1.661084],accel_mss,speed_ms,0,blend_radius_m)
  movel([0.085522, -0.803756, -2.776742, -1.131891, 1.570796, 1.656318],accel_mss,speed_ms,0,blend_radius_m)
  movel([0.080947, -0.808977, -2.775806, -1.127606, 1.570796, 1.651743],accel_mss,speed_ms,0,blend_radius_m)
  movel([0.076594, -0.814330, -2.774831, -1.123228, 1.570796, 1.647390],accel_mss,speed_ms,0,blend_radius_m)
  movel([0.072483, -0.819787, -2.773820, -1.118782, 1.570796, 1.643279],accel_mss,speed_ms,0,blend_radius_m)
  movel([0.068637, -0.825307, -2.772782, -1.114301, 1.570796, 1.639434],accel_mss,speed_ms,0,blend_radius_m)
  movel([0.065084, -0.830860, -2.771719, -1.109810, 1.570796, 1.635881],accel_mss,speed_ms,0,blend_radius_m)
  movel([0.065996, -0.829191, -2.772040, -1.111157, 1.570796, 1.636793],accel_mss,speed_ms,0,blend_radius_m)
  movel([0.066812, -0.827367, -2.772389, -1.112632, 1.570796, 1.637609],accel_mss,speed_ms,0,blend_radius_m)
  movel([0.068240, -0.823448, -2.773133, -1.115808, 1.570796, 1.639036],accel_mss,speed_ms,0,blend_radius_m)
  movel([0.070798, -0.815951, -2.774532, -1.121906, 1.570796, 1.641594],accel_mss,speed_ms,0,blend_radius_m)
  movel([0.073649, -0.809320, -2.775744, -1.127325, 1.570796, 1.644445],accel_mss,speed_ms,0,blend_radius_m)
  movel([0.076769, -0.802617, -2.776945, -1.132827, 1.570796, 1.647566],accel_mss,speed_ms,0,blend_radius_m)
  movel([0.080150, -0.795844, -2.778134, -1.138411, 1.570796, 1.650947],accel_mss,speed_ms,0,blend_radius_m)
  movel([0.083778, -0.789004, -2.779310, -1.144075, 1.570796, 1.654574],accel_mss,speed_ms,0,blend_radius_m)
  movel([0.087644, -0.782087, -2.780474, -1.149828, 1.570796, 1.658440],accel_mss,speed_ms,0,blend_radius_m)
  movel([0.091741, -0.775098, -2.781626, -1.155666, 1.570796, 1.662537],accel_mss,speed_ms,0,blend_radius_m)
  movel([0.100580, -0.760880, -2.783891, -1.167618, 1.570796, 1.671376],accel_mss,speed_ms,0,blend_radius_m)
  movel([0.096706, -0.765492, -2.783168, -1.163730, 1.570796, 1.667502],accel_mss,speed_ms,0,blend_radius_m)
  movel([0.084704, -0.778666, -2.781041, -1.152682, 1.570796, 1.655500],accel_mss,speed_ms,0,blend_radius_m)
  movel([0.080809, -0.783119, -2.780302, -1.148968, 1.570796, 1.651605],accel_mss,speed_ms,0,blend_radius_m)
  movel([0.077114, -0.787705, -2.779530, -1.145154, 1.570796, 1.647911],accel_mss,speed_ms,0,blend_radius_m)
  movel([0.073771, -0.792385, -2.778732, -1.141273, 1.570796, 1.644568],accel_mss,speed_ms,0,blend_radius_m)
  movel([0.070920, -0.797138, -2.777908, -1.137343, 1.570796, 1.641716],accel_mss,speed_ms,0,blend_radius_m)
  movel([0.074615, -0.789478, -2.779229, -1.143682, 1.570796, 1.645411],accel_mss,speed_ms,0,blend_radius_m)
  movel([0.078258, -0.781529, -2.780567, -1.150293, 1.570796, 1.649055],accel_mss,speed_ms,0,blend_radius_m)
  movel([0.082177, -0.773505, -2.781885, -1.157000, 1.570796, 1.652974],accel_mss,speed_ms,0,blend_radius_m)
  movel([0.084340, -0.769542, -2.782523, -1.160324, 1.570796, 1.655137],accel_mss,speed_ms,0,blend_radius_m)
  movel([0.086700, -0.765648, -2.783143, -1.163598, 1.570796, 1.657496],accel_mss,speed_ms,0,blend_radius_m)
  movel([0.095621, -0.752405, -2.785193, -1.174790, 1.570796, 1.666417],accel_mss,speed_ms,0,blend_radius_m)
  movel([0.104904, -0.738991, -2.787183, -1.186215, 1.570796, 1.675701],accel_mss,speed_ms,0,blend_radius_m)
  movel([0.097822, -0.746315, -2.786107, -1.179967, 1.570796, 1.668618],accel_mss,speed_ms,0,blend_radius_m)
  movel([0.091532, -0.753483, -2.785030, -1.173876, 1.570796, 1.662328],accel_mss,speed_ms,0,blend_radius_m)
  movel([0.085642, -0.760974, -2.783877, -1.167538, 1.570796, 1.656438],accel_mss,speed_ms,0,blend_radius_m)
  movel([0.079779, -0.769236, -2.782572, -1.160581, 1.570796, 1.650575],accel_mss,speed_ms,0,blend_radius_m)
  movel([0.082524, -0.764889, -2.783263, -1.164237, 1.570796, 1.653320],accel_mss,speed_ms,0,blend_radius_m)
  movel([0.084937, -0.760527, -2.783946, -1.167916, 1.570796, 1.655733],accel_mss,speed_ms,0,blend_radius_m)
  movel([0.093515, -0.742821, -2.786624, -1.182944, 1.570796, 1.664311],accel_mss,speed_ms,0,blend_radius_m)
  movel([0.095957, -0.738298, -2.787283, -1.186808, 1.570796, 1.666754],accel_mss,speed_ms,0,blend_radius_m)
  movel([0.098759, -0.733718, -2.787941, -1.190731, 1.570796, 1.669556],accel_mss,speed_ms,0,blend_radius_m)
  movel([0.102927, -0.727764, -2.788780, -1.195845, 1.570796, 1.673723],accel_mss,speed_ms,0,blend_radius_m)
  movel([0.106676, -0.723295, -2.789400, -1.199695, 1.570796, 1.677473],accel_mss,speed_ms,0,blend_radius_m)
  movel([0.107487, -0.722071, -2.789568, -1.200750, 1.570796, 1.678284],accel_mss,speed_ms,0,blend_radius_m)
  movel([0.107684, -0.721107, -2.789699, -1.201582, 1.570796, 1.678481],accel_mss,speed_ms,0,blend_radius_m)
  movel([0.107083, -0.721000, -2.789714, -1.201675, 1.570796, 1.677879],accel_mss,speed_ms,0,blend_radius_m)
  movel([0.105897, -0.721547, -2.789639, -1.201203, 1.570796, 1.676693],accel_mss,speed_ms,0,blend_radius_m)
  movel([0.104340, -0.722555, -2.789501, -1.200333, 1.570796, 1.675136],accel_mss,speed_ms,0,blend_radius_m)
  movel([0.100955, -0.725131, -2.789146, -1.198112, 1.570796, 1.671751],accel_mss,speed_ms,0,blend_radius_m)
  movel([0.098616, -0.727135, -2.788868, -1.196386, 1.570796, 1.669412],accel_mss,speed_ms,0,blend_radius_m)
  movel([0.101981, -0.721808, -2.789604, -1.200978, 1.570796, 1.672778],accel_mss,speed_ms,0,blend_radius_m)
  movel([0.106037, -0.716339, -2.790345, -1.205705, 1.570796, 1.676834],accel_mss,speed_ms,0,blend_radius_m)
  movel([0.114687, -0.705842, -2.791728, -1.214819, 1.570796, 1.685483],accel_mss,speed_ms,0,blend_radius_m)
  speed_ms = 0.005
  movel([0.114687, -0.699379, -2.785111, -1.227899, 1.570796, 1.685483],accel_mss,speed_ms,0,blend_radius_m)
  speed_ms = 0.040
  movel([0.097529, -0.710617, -2.783635, -1.218137, 1.570796, 1.668325],accel_mss,speed_ms,0,blend_radius_m)
  speed_ms = 0.005
  movel([0.097529, -0.717228, -2.790225, -1.204936, 1.570796, 1.668325],accel_mss,speed_ms,0,blend_radius_m)
  speed_ms = 0.025
  movel([0.095815, -0.716290, -2.790351, -1.205748, 1.570796, 1.666612],accel_mss,speed_ms,0,blend_radius_m)
  movel([0.093693, -0.716029, -2.790386, -1.205973, 1.570796, 1.664489],accel_mss,speed_ms,0,blend_radius_m)
  movel([0.091236, -0.716366, -2.790341, -1.205682, 1.570796, 1.662032],accel_mss,speed_ms,0,blend_radius_m)
  movel([0.088517, -0.717215, -2.790227, -1.204947, 1.570796, 1.659314],accel_mss,speed_ms,0,blend_radius_m)
  movel([0.085607, -0.718505, -2.790053, -1.203831, 1.570796, 1.656403],accel_mss,speed_ms,0,blend_radius_m)
  movel([0.082583, -0.720151, -2.789830, -1.202408, 1.570796, 1.653379],accel_mss,speed_ms,0,blend_radius_m)
  movel([0.076465, -0.724187, -2.789277, -1.198925, 1.570796, 1.647261],accel_mss,speed_ms,0,blend_radius_m)
  speed_ms = 0.005
  movel([0.076465, -0.717488, -2.782703, -1.212198, 1.570796, 1.647261],accel_mss,speed_ms,0,blend_radius_m)
  speed_ms = 0.040
  movel([0.100792, -0.695123, -2.785655, -1.231611, 1.570796, 1.671588],accel_mss,speed_ms,0,blend_radius_m)
  speed_ms = 0.005
  movel([0.100792, -0.701529, -2.792282, -1.218578, 1.570796, 1.671588],accel_mss,speed_ms,0,blend_radius_m)
  speed_ms = 0.025
  movel([0.099339, -0.698609, -2.792652, -1.221128, 1.570796, 1.670135],accel_mss,speed_ms,0,blend_radius_m)
  movel([0.097645, -0.696080, -2.792970, -1.223340, 1.570796, 1.668441],accel_mss,speed_ms,0,blend_radius_m)
  movel([0.095616, -0.694088, -2.793218, -1.225083, 1.570796, 1.666412],accel_mss,speed_ms,0,blend_radius_m)
  movel([0.093152, -0.692777, -2.793380, -1.226232, 1.570796, 1.663948],accel_mss,speed_ms,0,blend_radius_m)
  movel([0.090160, -0.692306, -2.793438, -1.226645, 1.570796, 1.660956],accel_mss,speed_ms,0,blend_radius_m)
  movel([0.086556, -0.692798, -2.793377, -1.226213, 1.570796, 1.657353],accel_mss,speed_ms,0,blend_radius_m)
  movel([0.082249, -0.694414, -2.793177, -1.224798, 1.570796, 1.653045],accel_mss,speed_ms,0,blend_radius_m)
  movel([0.079808, -0.695681, -2.793019, -1.223688, 1.570796, 1.650604],accel_mss,speed_ms,0,blend_radius_m)
  movel([0.077160, -0.697280, -2.792819, -1.222289, 1.570796, 1.647956],accel_mss,speed_ms,0,blend_radius_m)
  speed_ms = 0.005
  movel([0.077160, -0.690930, -2.786183, -1.235276, 1.570796, 1.647956],accel_mss,speed_ms,0,blend_radius_m)
  speed_ms = 0.040
  movel([0.097781, -0.672648, -2.788390, -1.251351, 1.570796, 1.668577],accel_mss,speed_ms,0,blend_radius_m)
  speed_ms = 0.005
  movel([0.097781, -0.678745, -2.795067, -1.238576, 1.570796, 1.668577],accel_mss,speed_ms,0,blend_radius_m)
  speed_ms = 0.025
  movel([0.096241, -0.671524, -2.795902, -1.244963, 1.570796, 1.667037],accel_mss,speed_ms,0,blend_radius_m)
  movel([0.095019, -0.668448, -2.796250, -1.247691, 1.570796, 1.665815],accel_mss,speed_ms,0,blend_radius_m)
  movel([0.093346, -0.665923, -2.796533, -1.249933, 1.570796, 1.664143],accel_mss,speed_ms,0,blend_radius_m)
  movel([0.091118, -0.664097, -2.796736, -1.251555, 1.570796, 1.661915],accel_mss,speed_ms,0,blend_radius_m)
  movel([0.088226, -0.663126, -2.796844, -1.252419, 1.570796, 1.659023],accel_mss,speed_ms,0,blend_radius_m)
  movel([0.084560, -0.663150, -2.796841, -1.252398, 1.570796, 1.655356],accel_mss,speed_ms,0,blend_radius_m)
  movel([0.080024, -0.664320, -2.796711, -1.251357, 1.570796, 1.650820],accel_mss,speed_ms,0,blend_radius_m)
  speed_ms = 0.005
  movel([0.080024, -0.658426, -2.790004, -1.263959, 1.570796, 1.650820],accel_mss,speed_ms,0,blend_radius_m)
  speed_ms = 0.040
  movel([0.099368, -0.648378, -2.791091, -1.272920, 1.570796, 1.670165],accel_mss,speed_ms,0,blend_radius_m)
  speed_ms = 0.005
  movel([0.099368, -0.654125, -2.797819, -1.260445, 1.570796, 1.670165],accel_mss,speed_ms,0,blend_radius_m)
  speed_ms = 0.025
  movel([0.099757, -0.648812, -2.798378, -1.265199, 1.570796, 1.670554],accel_mss,speed_ms,0,blend_radius_m)
  movel([0.099765, -0.643675, -2.798907, -1.269806, 1.570796, 1.670561],accel_mss,speed_ms,0,blend_radius_m)
  movel([0.099261, -0.638925, -2.799387, -1.274077, 1.570796, 1.670057],accel_mss,speed_ms,0,blend_radius_m)
  movel([0.098130, -0.634781, -2.799798, -1.277810, 1.570796, 1.668926],accel_mss,speed_ms,0,blend_radius_m)
  movel([0.096245, -0.631452, -2.800122, -1.280814, 1.570796, 1.667041],accel_mss,speed_ms,0,blend_radius_m)
  movel([0.094978, -0.630169, -2.800246, -1.281974, 1.570796, 1.665775],accel_mss,speed_ms,0,blend_radius_m)
  movel([0.091741, -0.628480, -2.800408, -1.283501, 1.570796, 1.662537],accel_mss,speed_ms,0,blend_radius_m)
  movel([0.089737, -0.628134, -2.800441, -1.283814, 1.570796, 1.660533],accel_mss,speed_ms,0,blend_radius_m)
  movel([0.087455, -0.628153, -2.800439, -1.283797, 1.570796, 1.658252],accel_mss,speed_ms,0,blend_radius_m)
  movel([0.084890, -0.628566, -2.800400, -1.283423, 1.570796, 1.655686],accel_mss,speed_ms,0,blend_radius_m)
  speed_ms = 0.005
  movel([0.084890, -0.623200, -2.793625, -1.295564, 1.570796, 1.655686],accel_mss,speed_ms,0,blend_radius_m)
  speed_ms = 0.040
  movel([0.105737, -0.611382, -2.794722, -1.306286, 1.570796, 1.676533],accel_mss,speed_ms,0,blend_radius_m)
  speed_ms = 0.005
  movel([0.105737, -0.616563, -2.801518, -1.294308, 1.570796, 1.676533],accel_mss,speed_ms,0,blend_radius_m)
  speed_ms = 0.025
  movel([0.106627, -0.610065, -2.802098, -1.300226, 1.570796, 1.677424],accel_mss,speed_ms,0,blend_radius_m)
  movel([0.106862, -0.603958, -2.802628, -1.305803, 1.570796, 1.677659],accel_mss,speed_ms,0,blend_radius_m)
  movel([0.106335, -0.598470, -2.803092, -1.310827, 1.570796, 1.677132],accel_mss,speed_ms,0,blend_radius_m)
  movel([0.104908, -0.593866, -2.803471, -1.315052, 1.570796, 1.675704],accel_mss,speed_ms,0,blend_radius_m)
  movel([0.102474, -0.590380, -2.803753, -1.318256, 1.570796, 1.673270],accel_mss,speed_ms,0,blend_radius_m)
  movel([0.100833, -0.589142, -2.803852, -1.319395, 1.570796, 1.671630],accel_mss,speed_ms,0,blend_radius_m)
  movel([0.098905, -0.588267, -2.803921, -1.320201, 1.570796, 1.669702],accel_mss,speed_ms,0,blend_radius_m)
  movel([0.096662, -0.587807, -2.803957, -1.320625, 1.570796, 1.667458],accel_mss,speed_ms,0,blend_radius_m)
  movel([0.094097, -0.587772, -2.803960, -1.320657, 1.570796, 1.664893],accel_mss,speed_ms,0,blend_radius_m)
  movel([0.091202, -0.588204, -2.803926, -1.320259, 1.570796, 1.661998],accel_mss,speed_ms,0,blend_radius_m)
  movel([0.087961, -0.589122, -2.803853, -1.319413, 1.570796, 1.658757],accel_mss,speed_ms,0,blend_radius_m)
  speed_ms = 0.005
  movel([0.087961, -0.584378, -2.797012, -1.330999, 1.570796, 1.658757],accel_mss,speed_ms,0,blend_radius_m)
  speed_ms = 0.040
  movel([-0.006407, -0.655979, -2.790273, -1.266137, 1.570796, 1.564389],accel_mss,speed_ms,0,blend_radius_m)
  speed_ms = 0.005
  movel([-0.006407, -0.661838, -2.796985, -1.253566, 1.570796, 1.564389],accel_mss,speed_ms,0,blend_radius_m)
  speed_ms = 0.025
  movel([-0.001379, -0.660923, -2.797085, -1.254380, 1.570796, 1.569417],accel_mss,speed_ms,0,blend_radius_m)
  movel([0.003243, -0.660752, -2.797104, -1.254532, 1.570796, 1.574039],accel_mss,speed_ms,0,blend_radius_m)
  movel([0.007469, -0.661277, -2.797047, -1.254066, 1.570796, 1.578265],accel_mss,speed_ms,0,blend_radius_m)
  movel([0.011300, -0.662449, -2.796918, -1.253022, 1.570796, 1.582096],accel_mss,speed_ms,0,blend_radius_m)
  movel([0.014728, -0.664229, -2.796722, -1.251439, 1.570796, 1.585525],accel_mss,speed_ms,0,blend_radius_m)
  movel([0.017776, -0.666557, -2.796463, -1.249369, 1.570796, 1.588572],accel_mss,speed_ms,0,blend_radius_m)
  movel([0.020434, -0.669400, -2.796143, -1.246846, 1.570796, 1.591230],accel_mss,speed_ms,0,blend_radius_m)
  movel([0.022726, -0.672687, -2.795769, -1.243933, 1.570796, 1.593522],accel_mss,speed_ms,0,blend_radius_m)
  movel([0.024647, -0.676382, -2.795343, -1.240664, 1.570796, 1.595443],accel_mss,speed_ms,0,blend_radius_m)
  movel([0.026223, -0.680423, -2.794870, -1.237095, 1.570796, 1.597019],accel_mss,speed_ms,0,blend_radius_m)
  movel([0.027455, -0.684761, -2.794355, -1.233273, 1.570796, 1.598251],accel_mss,speed_ms,0,blend_radius_m)
  movel([0.028360, -0.689351, -2.793800, -1.229238, 1.570796, 1.599156],accel_mss,speed_ms,0,blend_radius_m)
  movel([0.028950, -0.694126, -2.793213, -1.225050, 1.570796, 1.599746],accel_mss,speed_ms,0,blend_radius_m)
  movel([0.029231, -0.699058, -2.792596, -1.220735, 1.570796, 1.600028],accel_mss,speed_ms,0,blend_radius_m)
  movel([0.029222, -0.704076, -2.791956, -1.216356, 1.570796, 1.600018],accel_mss,speed_ms,0,blend_radius_m)
  movel([0.028939, -0.709141, -2.791299, -1.211949, 1.570796, 1.599735],accel_mss,speed_ms,0,blend_radius_m)
  movel([0.028205, -0.716074, -2.790380, -1.205934, 1.570796, 1.599001],accel_mss,speed_ms,0,blend_radius_m)
  movel([0.026905, -0.724269, -2.789265, -1.198855, 1.570796, 1.597702],accel_mss,speed_ms,0,blend_radius_m)
  movel([0.024855, -0.733170, -2.788019, -1.191201, 1.570796, 1.595652],accel_mss,speed_ms,0,blend_radius_m)
  movel([0.023495, -0.737715, -2.787367, -1.187307, 1.570796, 1.594291],accel_mss,speed_ms,0,blend_radius_m)
  movel([0.021889, -0.742224, -2.786711, -1.183454, 1.570796, 1.592685],accel_mss,speed_ms,0,blend_radius_m)
  movel([0.020001, -0.746649, -2.786058, -1.179682, 1.570796, 1.590797],accel_mss,speed_ms,0,blend_radius_m)
  movel([0.017822, -0.750906, -2.785420, -1.176063, 1.570796, 1.588618],accel_mss,speed_ms,0,blend_radius_m)
  movel([0.015318, -0.754948, -2.784807, -1.172635, 1.570796, 1.586114],accel_mss,speed_ms,0,blend_radius_m)
  movel([0.012467, -0.758714, -2.784227, -1.169447, 1.570796, 1.583264],accel_mss,speed_ms,0,blend_radius_m)
  movel([0.009250, -0.762134, -2.783695, -1.166559, 1.570796, 1.580047],accel_mss,speed_ms,0,blend_radius_m)
  movel([0.005635, -0.765165, -2.783219, -1.164005, 1.570796, 1.576431],accel_mss,speed_ms,0,blend_radius_m)
  movel([0.003664, -0.766516, -2.783005, -1.162867, 1.570796, 1.574460],accel_mss,speed_ms,0,blend_radius_m)
  movel([0.001583, -0.767751, -2.782809, -1.161829, 1.570796, 1.572379],accel_mss,speed_ms,0,blend_radius_m)
  movel([-0.002928, -0.769840, -2.782475, -1.160074, 1.570796, 1.567868],accel_mss,speed_ms,0,blend_radius_m)
  movel([-0.008186, -0.771618, -2.782190, -1.158582, 1.570796, 1.562610],accel_mss,speed_ms,0,blend_radius_m)
  movel([-0.013066, -0.772792, -2.782000, -1.157597, 1.570796, 1.557731],accel_mss,speed_ms,0,blend_radius_m)
  movel([-0.017616, -0.773436, -2.781896, -1.157057, 1.570796, 1.553180],accel_mss,speed_ms,0,blend_radius_m)
  movel([-0.021906, -0.773616, -2.781867, -1.156906, 1.570796, 1.548890],accel_mss,speed_ms,0,blend_radius_m)
  movel([-0.025984, -0.773394, -2.781902, -1.157092, 1.570796, 1.544813],accel_mss,speed_ms,0,blend_radius_m)
  movel([-0.029909, -0.772845, -2.781991, -1.157552, 1.570796, 1.540887],accel_mss,speed_ms,0,blend_radius_m)
  movel([-0.037530, -0.771021, -2.782286, -1.159083, 1.570796, 1.533266],accel_mss,speed_ms,0,blend_radius_m)
  movel([-0.045742, -0.768704, -2.782657, -1.161028, 1.570796, 1.525054],accel_mss,speed_ms,0,blend_radius_m)
  movel([-0.053769, -0.766215, -2.783053, -1.163121, 1.570796, 1.517027],accel_mss,speed_ms,0,blend_radius_m)
  movel([-0.061430, -0.763196, -2.783529, -1.165663, 1.570796, 1.509367],accel_mss,speed_ms,0,blend_radius_m)
  movel([-0.065060, -0.761365, -2.783816, -1.167208, 1.570796, 1.505736],accel_mss,speed_ms,0,blend_radius_m)
  movel([-0.068526, -0.759253, -2.784144, -1.168992, 1.570796, 1.502270],accel_mss,speed_ms,0,blend_radius_m)
  movel([-0.072951, -0.756765, -2.784528, -1.171096, 1.570796, 1.497845],accel_mss,speed_ms,0,blend_radius_m)
  movel([-0.077887, -0.754812, -2.784827, -1.172750, 1.570796, 1.492909],accel_mss,speed_ms,0,blend_radius_m)
  movel([-0.083253, -0.753354, -2.785049, -1.173985, 1.570796, 1.487543],accel_mss,speed_ms,0,blend_radius_m)
  movel([-0.088954, -0.752319, -2.785207, -1.174863, 1.570796, 1.481843],accel_mss,speed_ms,0,blend_radius_m)
  movel([-0.101008, -0.751309, -2.785359, -1.175721, 1.570796, 1.469788],accel_mss,speed_ms,0,blend_radius_m)
  movel([-0.113328, -0.751269, -2.785365, -1.175754, 1.570796, 1.457469],accel_mss,speed_ms,0,blend_radius_m)
  movel([-0.122964, -0.751974, -2.785259, -1.175156, 1.570796, 1.447833],accel_mss,speed_ms,0,blend_radius_m)
  movel([-0.133115, -0.753686, -2.784999, -1.173704, 1.570796, 1.437681],accel_mss,speed_ms,0,blend_radius_m)
  movel([-0.143727, -0.756412, -2.784582, -1.171395, 1.570796, 1.427070],accel_mss,speed_ms,0,blend_radius_m)
  movel([-0.154730, -0.760161, -2.784003, -1.168225, 1.570796, 1.416067],accel_mss,speed_ms,0,blend_radius_m)
  movel([-0.166061, -0.764920, -2.783258, -1.164211, 1.570796, 1.404735],accel_mss,speed_ms,0,blend_radius_m)
  movel([-0.171825, -0.767676, -2.782821, -1.161892, 1.570796, 1.398971],accel_mss,speed_ms,0,blend_radius_m)
  movel([-0.183512, -0.773930, -2.781816, -1.156643, 1.570796, 1.387285],accel_mss,speed_ms,0,blend_radius_m)
  movel([-0.189418, -0.777426, -2.781245, -1.153719, 1.570796, 1.381379],accel_mss,speed_ms,0,blend_radius_m)
  movel([-0.201295, -0.785130, -2.779965, -1.147294, 1.570796, 1.369501],accel_mss,speed_ms,0,blend_radius_m)
  movel([-0.209380, -0.790991, -2.778971, -1.142427, 1.570796, 1.361417],accel_mss,speed_ms,0,blend_radius_m)
  movel([-0.217381, -0.797420, -2.777859, -1.137110, 1.570796, 1.353415],accel_mss,speed_ms,0,blend_radius_m)
  movel([-0.225216, -0.804345, -2.776637, -1.131406, 1.570796, 1.345580],accel_mss,speed_ms,0,blend_radius_m)
  movel([-0.232807, -0.811710, -2.775310, -1.125369, 1.570796, 1.337990],accel_mss,speed_ms,0,blend_radius_m)
